{region 'Documentation'}
(*!
<summary>Capture once or compare against the retained snapshot after range validation.</summary>
*)
{endregion}
METHOD PROTECTED Assert
VAR
    ReferenceValue : REAL;
    ValuesEqual : BOOL;
    Value : REAL;
    InLowerIndex : DINT;
    InUpperIndex : DINT;
    MemoryLowerIndex : DINT;
    MemoryUpperIndex : DINT;
    MemoryEndIndex : LINT;
    EndIndex : LINT;
    Offset : LINT;
    InIndex : DINT;
    MemoryIndex : DINT;
    Message : STRING(GVL_Constants.MessageLength);
    ReferenceText : STRING(GVL_Constants.AssertionValueLength);
    ActualText : STRING(GVL_Constants.AssertionValueLength);
END_VAR
FEvaluationActive := ObservationActive AND FObservationPrevious AND FSnapshotValid;
FObservationPrevious := ObservationActive;

IF NOT ObservationActive THEN
    RETURN;
END_IF;

IF Result = E_Result.Error THEN
    RETURN;
END_IF;

// C0371: FB inputs are checked here before any reference access.
{warning disable C0371}
IF NOT __ISVALIDREF(IN) THEN
    Error(Message := 'Assertion error: IN reference is invalid.');
    RETURN;
END_IF;

IF NOT __ISVALIDREF(Memory) THEN
    Error(Message := 'Assertion error: Memory reference is invalid.');
    RETURN;
END_IF;

IF NOT Tc2_Utilities.RealIsFinite(x := Tolerance) THEN
    Error(Message := 'Assertion error: Tolerance must be finite.');
    RETURN;
END_IF;

IF Tolerance < 0.0 THEN
    Error(Message := 'Assertion error: Tolerance must not be negative.');
    RETURN;
END_IF;

InLowerIndex := LOWER_BOUND(IN, 1);
InUpperIndex := UPPER_BOUND(IN, 1);
MemoryLowerIndex := LOWER_BOUND(Memory, 1);
MemoryUpperIndex := UPPER_BOUND(Memory, 1);
EndIndex := DINT_TO_LINT(StartIndex) + USINT_TO_LINT(Length) - 1;
MemoryEndIndex := DINT_TO_LINT(MemoryLowerIndex) + USINT_TO_LINT(Length) - 1;

IF (Length = 0)
    OR (StartIndex < InLowerIndex) OR (StartIndex > InUpperIndex)
    OR (EndIndex > DINT_TO_LINT(InUpperIndex))
    OR (MemoryEndIndex > DINT_TO_LINT(MemoryUpperIndex)) THEN
    Message := CONCAT('Assertion error: array or memory range is invalid. StartIndex = ',
        DINT_TO_STRING(StartIndex));
    Message := CONCAT(Message, ', EndIndex = ');
    Message := CONCAT(Message, LINT_TO_STRING(EndIndex));
    Message := CONCAT(Message, ', Length = ');
    Message := CONCAT(Message, USINT_TO_STRING(Length));
    Message := CONCAT(Message, '.');
    Error(Message := Message);
    RETURN;
END_IF;

IF NOT FSnapshotValid THEN
    FOR Offset := 0 TO USINT_TO_LINT(Length) - 1 DO
        InIndex := LINT_TO_DINT(DINT_TO_LINT(StartIndex) + Offset);
        Value := IN[InIndex];
        IF Tc2_Utilities.RealIsNaN(x := Value) THEN
            Message := CONCAT('Assertion error: snapshot cannot contain NaN. IN index = ',
                DINT_TO_STRING(InIndex));
            Message := CONCAT(Message, '.');
            Error(Message := Message);
            RETURN;
        END_IF;
    END_FOR;
    FOR Offset := 0 TO USINT_TO_LINT(Length) - 1 DO
        InIndex := LINT_TO_DINT(DINT_TO_LINT(StartIndex) + Offset);
        MemoryIndex := LINT_TO_DINT(DINT_TO_LINT(MemoryLowerIndex) + Offset);
        Memory[MemoryIndex] := IN[InIndex];
    END_FOR;
    FSnapshotValid := TRUE;
    RETURN;
END_IF;

IF NOT EvaluationActive THEN
    RETURN;
END_IF;

IF Result = E_Result.Failed THEN
    RETURN;
END_IF;

FOR Offset := 0 TO USINT_TO_LINT(Length) - 1 DO
    InIndex := LINT_TO_DINT(DINT_TO_LINT(StartIndex) + Offset);
    MemoryIndex := LINT_TO_DINT(DINT_TO_LINT(MemoryLowerIndex) + Offset);
    Value := IN[InIndex];
    ReferenceValue := Memory[MemoryIndex];
    ValuesEqual := FALSE;
    IF NOT Tc2_Utilities.RealIsNaN(x := Value) THEN
        IF Value = ReferenceValue THEN
            ValuesEqual := TRUE;
        ELSIF Tc2_Utilities.RealIsFinite(x := Value)
            AND Tc2_Utilities.RealIsFinite(x := ReferenceValue) THEN
            ValuesEqual := IsWithinTolerance_Real(IN := Value,
                Expected := ReferenceValue,
                Tolerance := Tolerance);
        END_IF;
    END_IF;
    IF NOT ValuesEqual THEN
        Value := Memory[MemoryIndex];
        IF Tc2_Utilities.RealIsFinite(x := Value) THEN
            ReferenceText := CreateAssertionTextValue_Real(Value := Value);
        ELSE
            ReferenceText := '<non-finite>';
        END_IF;
        Value := IN[InIndex];
        IF Tc2_Utilities.RealIsFinite(x := Value) THEN
            ActualText := CreateAssertionTextValue_Real(Value := IN[InIndex]);
        ELSE
            ActualText := '<non-finite>';
        END_IF;
        Message := CONCAT('Assertion failed: array value changed. Reference[',
            DINT_TO_STRING(MemoryIndex));
        Message := CONCAT(Message, '] = ');
        Message := CONCAT(Message, ReferenceText);
        Message := CONCAT(Message, ', IN[');
        Message := CONCAT(Message, DINT_TO_STRING(InIndex));
        Message := CONCAT(Message, '] = ');
        Message := CONCAT(Message, ActualText);
        Message := CONCAT(Message, '.');
        Message := CONCAT(Message, ' Tolerance = ');
        Message := CONCAT(Message, CreateAssertionTextValue_Real(Value := Tolerance));
        Fail(Message := Message);
        RETURN;
    END_IF;
END_FOR;

Pass();
{warning restore C0371}
END_METHOD

{region 'Documentation'}
(*!
<summary>Current/last call has consecutive observation and an existing snapshot.</summary>
*)
{endregion}
{attribute 'monitoring' := 'call'}
PROPERTY PUBLIC EvaluationActive : BOOL //! Current/last call has consecutive observation and an existing snapshot.
GET // PUBLIC
EvaluationActive := FEvaluationActive;
END_GET
END_PROPERTY

{region 'Documentation'}
(*!
<summary>Invalidate the snapshot and observation history.</summary>
<description>

Does not clear external Memory. The next active observation captures a new snapshot
before comparison.

</description>
*)
{endregion}
METHOD PROTECTED ResetAssertion
FSnapshotValid := FALSE;
FObservationPrevious := FALSE;
FEvaluationActive := FALSE;
END_METHOD

END_FUNCTION_BLOCK

// ---- Framework/Assertions/POU/Utilities/IsWithinTolerance_Real.TcPOU
{region 'Documentation'}
(*!
<summary>Tests absolute tolerance without overflowing the typed difference. Requires finite inputs and a finite, non-negative tolerance; the caller validates them.</summary>
*)
{endregion}
FUNCTION INTERNAL IsWithinTolerance_Real : BOOL //! TRUE when the absolute difference is within Tolerance; caller must supply finite valid inputs.
VAR_INPUT
    IN : REAL; //! Actual value checked or observed by this Assertion.
    Expected : REAL; //! Reference value for comparison with IN.
    Tolerance : REAL; //! Maximum absolute difference accepted as equal; must be finite and non-negative.
END_VAR
VAR
    ActualMagnitude : REAL;
    ExpectedMagnitude : REAL;
    LargeMagnitude : REAL;
    SmallMagnitude : REAL;
    RemainingMagnitude : REAL;
    Difference : REAL;
END_VAR
VAR CONSTANT
    MaxFinite : REAL := REAL#3.40282346638528859811704183484516925440E38;
    HalfMaxFinite : REAL := MaxFinite / REAL#2.0;
END_VAR

IsWithinTolerance_Real := FALSE;

IF ((IN < 0.0) AND (Expected > 0.0)) OR ((IN > 0.0) AND (Expected < 0.0)) THEN
    ActualMagnitude := ABS(IN);
    ExpectedMagnitude := ABS(Expected);
    LargeMagnitude := MAX(ActualMagnitude, ExpectedMagnitude);
    SmallMagnitude := MIN(ActualMagnitude, ExpectedMagnitude);

    IF LargeMagnitude >= HalfMaxFinite THEN
        // Exact subtraction: MaxFinite and LargeMagnitude are within a factor of two.
        RemainingMagnitude := MaxFinite - LargeMagnitude;
        IF SmallMagnitude > RemainingMagnitude THEN
            RETURN;
        END_IF;
    END_IF;
END_IF;

Difference := ABS(IN - Expected);
IsWithinTolerance_Real := Difference <= Tolerance;

END_FUNCTION

// ---- Framework/Assertions/POU/Arrays/LReal/AssertArrayNoValueChange_LReal.TcPOU
{region 'Documentation'}
(*!
<summary>Captures one snapshot until Reset; Disable/Re-Enable never replaces it.</summary>
<description>

Disabling observation preserves the original snapshot. Re-enabling requires a fresh
preceding observation before comparisons resume; it does not replace that snapshot.

StartIndex is an absolute IN index and Length selects 1..255 elements within IN. Memory
must have at least Length elements from its own lower bound. Invalid references or ranges
report Error.

The caller provides dedicated writable Memory that must not overlap IN; overlap is not
checked. Keep bindings, selected range and snapshot contents stable until Reset. Reset
invalidates the snapshot without clearing Memory bytes.

Snapshot capture rejects NaN with Error but accepts either infinity. Later NaN is a
mismatch; equal signed infinities match.

Tolerance is absolute, in the same units as the values, finite and non-negative. Its
default zero requests exact comparison. The equality boundary is inclusive; larger differences
are unequal. Difference checking avoids overflow for large finite operands.

Numeric diagnostics use the formatter's default six significant digits; rounding affects
the message only, not the comparison.

</description>
*)
{endregion}
FUNCTION_BLOCK AssertArrayNoValueChange_LReal EXTENDS AssertionBase
VAR_INPUT
    Tolerance : LREAL := 0.0; //! Maximum absolute allowed difference; finite and non-negative.
    StartIndex : DINT; //! First selected index in IN; uses the array's declared index range, not a zero-based offset.
    Length : USINT; //! Number of monitored elements, from 1 through 255.
END_VAR
VAR_IN_OUT CONSTANT
    IN : ARRAY[*] OF LREAL; //! Read-only actual data; the selected range must remain stable during the call.
END_VAR
VAR_IN_OUT
    Memory : ARRAY[*] OF LREAL; //! Dedicated snapshot storage; only this assertion writes its selected elements.
END_VAR
VAR
    FSnapshotValid : BOOL;
    FObservationPrevious : BOOL;
    FEvaluationActive : BOOL;
END_VAR

SUPER^();

{region 'Documentation'}
(*!
<summary>Capture once or compare against the retained snapshot after range validation.</summary>
*)
{endregion}
METHOD PROTECTED Assert
VAR
    ReferenceValue : LREAL;
    ValuesEqual : BOOL;
    Value : LREAL;
    InLowerIndex : DINT;
    InUpperIndex : DINT;
    MemoryLowerIndex : DINT;
    MemoryUpperIndex : DINT;
    MemoryEndIndex : LINT;
    EndIndex : LINT;
    Offset : LINT;
    InIndex : DINT;
    MemoryIndex : DINT;
    Message : STRING(GVL_Constants.MessageLength);
    ReferenceText : STRING(GVL_Constants.AssertionValueLength);
    ActualText : STRING(GVL_Constants.AssertionValueLength);
END_VAR
FEvaluationActive := ObservationActive AND FObservationPrevious AND FSnapshotValid;
FObservationPrevious := ObservationActive;

IF NOT ObservationActive THEN
    RETURN;
END_IF;

IF Result = E_Result.Error THEN
    RETURN;
END_IF;

// C0371: FB inputs are checked here before any reference access.
{warning disable C0371}
IF NOT __ISVALIDREF(IN) THEN
    Error(Message := 'Assertion error: IN reference is invalid.');
    RETURN;
END_IF;

IF NOT __ISVALIDREF(Memory) THEN
    Error(Message := 'Assertion error: Memory reference is invalid.');
    RETURN;
END_IF;

IF NOT Tc2_Utilities.LrealIsFinite(x := Tolerance) THEN
    Error(Message := 'Assertion error: Tolerance must be finite.');
    RETURN;
END_IF;

IF Tolerance < 0.0 THEN
    Error(Message := 'Assertion error: Tolerance must not be negative.');
    RETURN;
END_IF;

InLowerIndex := LOWER_BOUND(IN, 1);
InUpperIndex := UPPER_BOUND(IN, 1);
MemoryLowerIndex := LOWER_BOUND(Memory, 1);
MemoryUpperIndex := UPPER_BOUND(Memory, 1);
EndIndex := DINT_TO_LINT(StartIndex) + USINT_TO_LINT(Length) - 1;
MemoryEndIndex := DINT_TO_LINT(MemoryLowerIndex) + USINT_TO_LINT(Length) - 1;

IF (Length = 0)
    OR (StartIndex < InLowerIndex) OR (StartIndex > InUpperIndex)
    OR (EndIndex > DINT_TO_LINT(InUpperIndex))
    OR (MemoryEndIndex > DINT_TO_LINT(MemoryUpperIndex)) THEN
    Message := CONCAT('Assertion error: array or memory range is invalid. StartIndex = ',
        DINT_TO_STRING(StartIndex));
    Message := CONCAT(Message, ', EndIndex = ');
    Message := CONCAT(Message, LINT_TO_STRING(EndIndex));
    Message := CONCAT(Message, ', Length = ');
    Message := CONCAT(Message, USINT_TO_STRING(Length));
    Message := CONCAT(Message, '.');
    Error(Message := Message);
    RETURN;
END_IF;

IF NOT FSnapshotValid THEN
    FOR Offset := 0 TO USINT_TO_LINT(Length) - 1 DO
        InIndex := LINT_TO_DINT(DINT_TO_LINT(StartIndex) + Offset);
        Value := IN[InIndex];
        IF Tc2_Utilities.LrealIsNaN(x := Value) THEN
            Message := CONCAT('Assertion error: snapshot cannot contain NaN. IN index = ',
                DINT_TO_STRING(InIndex));
            Message := CONCAT(Message, '.');
            Error(Message := Message);
            RETURN;
        END_IF;
    END_FOR;
    FOR Offset := 0 TO USINT_TO_LINT(Length) - 1 DO
        InIndex := LINT_TO_DINT(DINT_TO_LINT(StartIndex) + Offset);
        MemoryIndex := LINT_TO_DINT(DINT_TO_LINT(MemoryLowerIndex) + Offset);
        Memory[MemoryIndex] := IN[InIndex];
    END_FOR;
    FSnapshotValid := TRUE;
    RETURN;
END_IF;

IF NOT EvaluationActive THEN
    RETURN;
END_IF;

IF Result = E_Result.Failed THEN
    RETURN;
END_IF;

FOR Offset := 0 TO USINT_TO_LINT(Length) - 1 DO
    InIndex := LINT_TO_DINT(DINT_TO_LINT(StartIndex) + Offset);
    MemoryIndex := LINT_TO_DINT(DINT_TO_LINT(MemoryLowerIndex) + Offset);
    Value := IN[InIndex];
    ReferenceValue := Memory[MemoryIndex];
    ValuesEqual := FALSE;
    IF NOT Tc2_Utilities.LrealIsNaN(x := Value) THEN
        IF Value = ReferenceValue THEN
            ValuesEqual := TRUE;
        ELSIF Tc2_Utilities.LrealIsFinite(x := Value)
            AND Tc2_Utilities.LrealIsFinite(x := ReferenceValue) THEN
            ValuesEqual := IsWithinTolerance_LReal(IN := Value,
                Expected := ReferenceValue,
                Tolerance := Tolerance);
        END_IF;
    END_IF;
    IF NOT ValuesEqual THEN
        Value := Memory[MemoryIndex];
        IF Tc2_Utilities.LrealIsFinite(x := Value) THEN
            ReferenceText := CreateAssertionTextValue_LReal(Value := Value);
        ELSE
            ReferenceText := '<non-finite>';
        END_IF;
        Value := IN[InIndex];
        IF Tc2_Utilities.LrealIsFinite(x := Value) THEN
            ActualText := CreateAssertionTextValue_LReal(Value := IN[InIndex]);
        ELSE
            ActualText := '<non-finite>';
        END_IF;
        Message := CONCAT('Assertion failed: array value changed. Reference[',
            DINT_TO_STRING(MemoryIndex));
        Message := CONCAT(Message, '] = ');
        Message := CONCAT(Message, ReferenceText);
        Message := CONCAT(Message, ', IN[');
        Message := CONCAT(Message, DINT_TO_STRING(InIndex));
        Message := CONCAT(Message, '] = ');
        Message := CONCAT(Message, ActualText);
        Message := CONCAT(Message, '.');
        Message := CONCAT(Message, ' Tolerance = ');
        Message := CONCAT(Message, CreateAssertionTextValue_LReal(Value := Tolerance));
        Fail(Message := Message);
        RETURN;
    END_IF;
END_FOR;

Pass();
{warning restore C0371}
END_METHOD

{region 'Documentation'}
(*!
<summary>Current/last call has consecutive observation and an existing snapshot.</summary>
*)
{endregion}
{attribute 'monitoring' := 'call'}
PROPERTY PUBLIC EvaluationActive : BOOL //! Current/last call has consecutive observation and an existing snapshot.
GET // PUBLIC
EvaluationActive := FEvaluationActive;
END_GET
END_PROPERTY

{region 'Documentation'}
(*!
<summary>Invalidate the snapshot and observation history.</summary>
<description>

Does not clear external Memory. The next active observation captures a new snapshot
before comparison.

</description>
*)
{endregion}
METHOD PROTECTED ResetAssertion
FSnapshotValid := FALSE;
FObservationPrevious := FALSE;
FEvaluationActive := FALSE;
END_METHOD

END_FUNCTION_BLOCK

// ---- SelfTests/TestSuites/TestSuite_AssertionText.TcPOU
{region 'Documentation'}
(*!
<summary>Checks text, token and diagnostic boundaries with isolated Assertion subjects.</summary>
*)
{endregion}
FUNCTION_BLOCK TestSuite_AssertionText EXTENDS TestSuiteBase
VAR
    FTextComparison : Test_AssertionTextComparison;
    FTextSearch : Test_AssertionTextSearch;
    FTextDiagnostics : Test_AssertionTextDiagnostics;
    FValueTokenCount : Test_AssertionValueTokenCount;
    FArrayTokenCount : Test_AssertionArrayTokenCount;
    FLengthUntil : Test_AssertionLengthUntil;
    FTestCases : ARRAY[1..TestCaseCapacity] OF I_TestCase;
END_VAR
VAR CONSTANT
    TestCaseCapacity : UINT := 6;
END_VAR

SUPER^();

{region 'Documentation'}
(*!
<summary>Initializes six isolated text and token Test Cases and registers them serially.</summary>
*)
{endregion}
METHOD PROTECTED Configure
VAR_IN_OUT
    // SA0167: Borrowed owner builder; no temporary instance is created.
    {attribute 'analysis' := '-167'}
    Builder : TestSuiteConfigurationBuilder; //! Borrowed owner configuration builder used only during this Configure call; register this owner's concrete children.
END_VAR
VAR
    TestConfig : ST_TestCaseConfig;
END_VAR
Builder.Initialize(Mode := E_OrchestrationMode.Serial,
    TestCases := FTestCases);
FTextComparison.Initialize(Parent := THIS^,
    TestName := 'TextComparison',
    Config := TestConfig);
Builder.Register(TestCase := FTextComparison);
FTextSearch.Initialize(Parent := THIS^,
    TestName := 'TextSearch',
    Config := TestConfig);
Builder.Register(TestCase := FTextSearch);
FTextDiagnostics.Initialize(Parent := THIS^,
    TestName := 'TextDiagnostics',
    Config := TestConfig);
Builder.Register(TestCase := FTextDiagnostics);
FValueTokenCount.Initialize(Parent := THIS^,
    TestName := 'ValueTokenCount',
    Config := TestConfig);
Builder.Register(TestCase := FValueTokenCount);
FArrayTokenCount.Initialize(Parent := THIS^,
    TestName := 'ArrayTokenCount',
    Config := TestConfig);
Builder.Register(TestCase := FArrayTokenCount);
FLengthUntil.Initialize(Parent := THIS^,
    TestName := 'LengthUntil',
    Config := TestConfig);
Builder.Register(TestCase := FLengthUntil);
END_METHOD

{region 'Documentation'}
(*!
<summary>Returns a registered scenario using its original array index.</summary>
*)
{endregion}
METHOD PUBLIC GetTestCase : I_TestCase //! Typed child interface at the original array index; zero when no entry is available.
VAR_INPUT
    Index : DINT; //! Original occupied child-array index, rather than an ordinal position.
END_VAR
GetTestCase := 0;
IF (ChildCount = 0) OR (Index < ChildArrayLowerBound)
    OR (DINT_TO_LINT(Index) >= DINT_TO_LINT(ChildArrayLowerBound) + UINT_TO_LINT(ChildCount)) THEN
    RETURN;
END_IF;
GetTestCase := FTestCases[Index];
END_METHOD

{region 'Documentation'}
(*!
<summary>Calls every owned scenario once per initialized Suite cycle.</summary>
*)
{endregion}
METHOD PROTECTED ProcessTestCases
FTextComparison();
FTextSearch();
FTextDiagnostics();
FValueTokenCount();
FArrayTokenCount();
FLengthUntil();
END_METHOD

END_FUNCTION_BLOCK

// ---- SelfTests/TestCases/TestSuite_AssertionText/Test_AssertionTextComparison.TcPOU
{region 'Documentation'}
(*!
<summary>Checks exact STRING/WSTRING comparisons and configured length boundaries.</summary>
<description>
Equality and inequality share explicit operands, but each result is asserted.
Wide-code-unit cases distinguish a zero low byte from the WSTRING terminator
and equal low bytes from equal code units. Capacity tests use the configured
content limits, including the last character and one excessive character.
Each scenario occupies two calls: Reset with valid bindings, then evaluation.
ProcessAssertions checks each call before ProcessTests advances. Literal expected
results belong to SelectScenario, not to a copy of the production comparison.
The local capture is cleared before each call and checked in subject-call order.
FirstFailedScenario and FailedDuringEvaluation retain the first mismatch.
Caller text buffers provide at least one extra character of capacity so overlength tests
reach the real read-only reference API without an intermediate truncating copy.
</description>
*)
{endregion}
FUNCTION_BLOCK Test_AssertionTextComparison EXTENDS TestCaseBase
VAR
    FEqual : AssertEqual_String;
    FEqualExpectedResult : E_Result;
    FNotEqual : AssertNotEqual_String;
    FNotEqualExpectedResult : E_Result;
    FWideEqual : AssertEqual_WString;
    FWideEqualExpectedResult : E_Result;
    FWideNotEqual : AssertNotEqual_WString;
    FWideNotEqualExpectedResult : E_Result;
    FInput : STRING(InputCapacity);
    FInputBefore : STRING(InputCapacity);
    FWideInput : WSTRING(WideInputCapacity);
    FWideInputBefore : WSTRING(WideInputCapacity);
    FExpected : STRING(InputCapacity);
    FExpectedBefore : STRING(InputCapacity);
    FWideExpected : WSTRING(WideInputCapacity);
    FWideExpectedBefore : WSTRING(WideInputCapacity);
    FCapture : EventBuffer;
    FEvents : ARRAY[1..CaptureLength] OF ST_Event;
    FCaptureFifo : ST_FifoStatus;
    FCaptureStatus : ST_EventBufferStatus;
    FSetupValid : BOOL;
    FScenario : UINT;
    FChecked : BOOL;
    FEvaluateSubjects : BOOL;
    FObservationReady : BOOL;
    FFirstFailedScenario : UINT;
    FFailedDuringEvaluation : BOOL;
    FResultsMatch : BOOL;
    FResults : AssertTrue;
    FActivityMatch : BOOL;
    FActivity : AssertTrue;
    FInputsMatch : BOOL;
    FInputs : AssertTrue;
    FFindingsMatch : BOOL;
    FFindings : AssertTrue;
END_VAR
VAR CONSTANT
    InputCapacity : UINT := Param_Assertions.AssertionStringLength + 1;
    // XAE rejects a computed WSTRING capacity here. Covers the default limit plus one.
    // CheckInitialization rejects a configuration exceeding this test storage.
    WideInputCapacity : UINT := 81;
    CaptureLength : UINT := 8;
    ScenarioExact : UINT := 1;
    ScenarioEmpty : UINT := 2;
    ScenarioCaseSensitive : UINT := 3;
    ScenarioFirstCharacter : UINT := 4;
    ScenarioLastCharacter : UINT := 5;
    ScenarioDifferentLength : UINT := 6;
    ScenarioWideHighByte : UINT := 7;
    ScenarioWideZeroLowByte : UINT := 8;
    ScenarioBelowCapacity : UINT := 9;
    ScenarioAtCapacity : UINT := 10;
    ScenarioLastAtCapacity : UINT := 11;
    ScenarioInputOverCapacity : UINT := 12;
    ScenarioExpectedOverCapacity : UINT := 13;
    LastScenario : UINT := ScenarioExpectedOverCapacity;
END_VAR

SUPER^();

{region 'Documentation'}
(*!
<summary>Aggregates only outer checks, not intentionally failing subjects.</summary>
*)
{endregion}
METHOD PROTECTED AggregateResults
VAR_INPUT
    Aggregator : I_ResultAggregator; //! Borrowed result sink owned by the outer Test Case; add this test's checking Assertions without resetting or retaining the sink.
END_VAR
Aggregator.AddProvider(Provider := FResults);
Aggregator.AddProvider(Provider := FActivity);
Aggregator.AddProvider(Provider := FInputs);
Aggregator.AddProvider(Provider := FFindings);
END_METHOD

{region 'Documentation'}
(*!
<summary>Calls each inherited production subject once with caller-owned text storage.</summary>
*)
{endregion}
METHOD PRIVATE CallSubjects
FEqual(Enable := TRUE,
    State := E_State.Running,
    IN := FInput,
    Expected := FExpected);
FNotEqual(Enable := TRUE,
    State := E_State.Running,
    IN := FInput,
    Expected := FExpected);
FWideEqual(Enable := TRUE,
    State := E_State.Running,
    IN := FWideInput,
    Expected := FWideExpected);
FWideNotEqual(Enable := TRUE,
    State := E_State.Running,
    IN := FWideInput,
    Expected := FWideExpected);
END_METHOD

{region 'Documentation'}
(*!
<summary>Checks one subject finding in call order; expected outcomes come from the scenario.</summary>
*)
{endregion}
METHOD PRIVATE CheckFinding : BOOL //! TRUE when the required finding checks pass; calls requiring no finding also succeed.
VAR_INPUT
    Subject : I_Assertion; //! Assertion interface supplying the expected finding identity.
    ExpectedResult : E_Result; //! Independently authored result expected in the captured finding.
END_VAR
VAR_IN_OUT
    Index : UINT; //! One-based next finding index; advanced when this call checks a required finding.
END_VAR
CheckFinding := TRUE;
IF FEvaluateSubjects AND ((ExpectedResult = E_Result.Failed)
    OR (ExpectedResult = E_Result.Error)) THEN
    CheckFinding := (FEvents[Index].SequenceId = UINT_TO_UDINT(Index))
        AND (FEvents[Index].Name = Subject.Name)
        AND (FEvents[Index].OwnerScope = E_OwnerScope.Assertion)
        AND (FEvents[Index].EventType = E_EventType.Result)
        AND (FEvents[Index].State = E_State.Running)
        AND (FEvents[Index].Result = ExpectedResult)
        AND (FEvents[Index].Message <> '');
    Index := Index + 1;
END_IF;
END_METHOD

{region 'Documentation'}
(*!
<summary>Checks exact finding count and identities; at most one finding per subject.</summary>
*)
{endregion}
METHOD PRIVATE CheckFindings
VAR
    Index : UINT;
    Matches : BOOL;
END_VAR
Index := 1;
FFindingsMatch := TRUE;
Matches := CheckFinding(Subject := FEqual,
    ExpectedResult := FEqualExpectedResult,
    Index := Index);
FFindingsMatch := FFindingsMatch AND Matches;
Matches := CheckFinding(Subject := FNotEqual,
    ExpectedResult := FNotEqualExpectedResult,
    Index := Index);
FFindingsMatch := FFindingsMatch AND Matches;
Matches := CheckFinding(Subject := FWideEqual,
    ExpectedResult := FWideEqualExpectedResult,
    Index := Index);
FFindingsMatch := FFindingsMatch AND Matches;
Matches := CheckFinding(Subject := FWideNotEqual,
    ExpectedResult := FWideNotEqualExpectedResult,
    Index := Index);
FFindingsMatch := FFindingsMatch AND Matches;
FFindingsMatch := FFindingsMatch
    AND (FCaptureStatus.SequenceId = UINT_TO_UDINT(Index - 1))
    AND (FCaptureStatus.LostEventCount = 0);
END_METHOD

{region 'Documentation'}
(*!
<summary>Rejects incomplete subject, capture or outer Assertion setup.</summary>
*)
{endregion}
METHOD PROTECTED CheckInitialization : BOOL //! TRUE when the inherited initialization check and this concrete fixture check both accept the setup.
CheckInitialization := SUPER^.CheckInitialization();
IF NOT CheckInitialization THEN
    RETURN;
END_IF;

CheckInitialization := FSetupValid
    AND (Param_Assertions.AssertionStringLength >= 5)
    AND (Param_Assertions.AssertionWStringLength >= 5)
    AND (Param_Assertions.AssertionWStringLength < WideInputCapacity)
    AND FResults.IsInitialized
    AND FActivity.IsInitialized
    AND FInputs.IsInitialized
    AND FFindings.IsInitialized;
IF NOT CheckInitialization THEN
    EventPublisher.PublishEvent(Event := CreateFrameworkEvent(Name := Name,
        ResourceName := '',
        State := State,
        Severity := E_EventSeverity.Error,
        Message := 'Text selftest setup failed.'));
END_IF;
END_METHOD

{region 'Documentation'}
(*!
<summary>Checks literal evaluation results, or NotEvaluated on the reset call.</summary>
*)
{endregion}
METHOD PRIVATE CheckResults
IF FEvaluateSubjects THEN
    FResultsMatch := (FEqual.Result = FEqualExpectedResult)
        AND (FNotEqual.Result = FNotEqualExpectedResult)
        AND (FWideEqual.Result = FWideEqualExpectedResult)
        AND (FWideNotEqual.Result = FWideNotEqualExpectedResult);
ELSE
    FResultsMatch := (FEqual.Result = E_Result.NotEvaluated)
        AND (FNotEqual.Result = E_Result.NotEvaluated)
        AND (FWideEqual.Result = E_Result.NotEvaluated)
        AND (FWideNotEqual.Result = E_Result.NotEvaluated);
END_IF;
FActivityMatch := FEqual.Enabled
    AND (FEqual.ObservationActive = FEvaluateSubjects)
    AND (FEqual.EvaluationActive = FEvaluateSubjects)
    AND FNotEqual.Enabled
    AND (FNotEqual.ObservationActive = FEvaluateSubjects)
    AND (FNotEqual.EvaluationActive = FEvaluateSubjects)
    AND FWideEqual.Enabled
    AND (FWideEqual.ObservationActive = FEvaluateSubjects)
    AND (FWideEqual.EvaluationActive = FEvaluateSubjects)
    AND FWideNotEqual.Enabled
    AND (FWideNotEqual.ObservationActive = FEvaluateSubjects)
    AND (FWideNotEqual.EvaluationActive = FEvaluateSubjects);
END_METHOD

{region 'Documentation'}
(*!
<summary>Initializes outer checks and isolates intentional subject findings.</summary>
*)
{endregion}
METHOD PROTECTED Configure
VAR
    Initialized : BOOL;
END_VAR
FPreparationStateCount := 0;
FTestStateCount := 1;
FResults.Initialize(Parent := THIS^,
    AssertionName := 'Results');
FActivity.Initialize(Parent := THIS^,
    AssertionName := 'Activity');
FInputs.Initialize(Parent := THIS^,
    AssertionName := 'Inputs');
FFindings.Initialize(Parent := THIS^,
    AssertionName := 'Findings');
FSetupValid := FCapture.Initialize(Buffer := FEvents,
    FifoControl := FCaptureFifo,
    Status := FCaptureStatus);
FEqual.BindPublisher(Publisher := FCapture);
Initialized := FEqual.Initialize(Parent := THIS^,
    AssertionName := 'Equal');
FSetupValid := FSetupValid AND Initialized;
FNotEqual.BindPublisher(Publisher := FCapture);
Initialized := FNotEqual.Initialize(Parent := THIS^,
    AssertionName := 'NotEqual');
FSetupValid := FSetupValid AND Initialized;
FWideEqual.BindPublisher(Publisher := FCapture);
Initialized := FWideEqual.Initialize(Parent := THIS^,
    AssertionName := 'WideEqual');
FSetupValid := FSetupValid AND Initialized;
FWideNotEqual.BindPublisher(Publisher := FCapture);
Initialized := FWideNotEqual.Initialize(Parent := THIS^,
    AssertionName := 'WideNotEqual');
FSetupValid := FSetupValid AND Initialized;
END_METHOD

{region 'Documentation'}
(*!
<summary>Completes abort; no asynchronous resource is owned.</summary>
*)
{endregion}
METHOD PROTECTED ProcessAbort
VAR_INPUT
    Enable : BOOL; //! Phase permission supplied by the owning Test Case; FALSE does not authorize progression, while observation may continue.
END_VAR
IF Enable THEN
    CompleteAbort();
END_IF;
END_METHOD

{region 'Documentation'}
(*!
<summary>Latches this call's checks before progression is permitted.</summary>
*)
{endregion}
METHOD PROTECTED ProcessAssertions
VAR_INPUT
    Enable : BOOL; //! Phase permission supplied by the owning Test Case; FALSE does not authorize progression, while observation may continue.
END_VAR
VAR
    Check : BOOL;
END_VAR
Check := Enable AND FObservationReady;
FResults(Enable := Check,
    State := State,
    IN := FResultsMatch);
FActivity(Enable := Check,
    State := State,
    IN := FActivityMatch);
FInputs(Enable := Check,
    State := State,
    IN := FInputsMatch);
FFindings(Enable := Check,
    State := State,
    IN := FFindingsMatch);
IF Check THEN
    FChecked := TRUE;
END_IF;
END_METHOD

{region 'Documentation'}
(*!
<summary>No Preparation phase is needed.</summary>
*)
{endregion}
METHOD PROTECTED ProcessPreparations
VAR_INPUT
    // SA0033: Required hook; this test has no Preparation phase.
    {attribute 'analysis' := '-33'}
    Enable : BOOL; //! Phase permission supplied by the owning Test Case; FALSE does not authorize progression, while observation may continue.
END_VAR
END_METHOD

{region 'Documentation'}
(*!
<summary>Restarts the scenario sequence and outer checks.</summary>
*)
{endregion}
METHOD PROTECTED ProcessReset
FScenario := ScenarioExact;
FChecked := FALSE;
FEvaluateSubjects := FALSE;
FObservationReady := FALSE;
FFirstFailedScenario := 0;
FFailedDuringEvaluation := FALSE;
FCapture.Reset();
ResetSubjects();
FResults.Reset();
FActivity.Reset();
FInputs.Reset();
FFindings.Reset();
CompleteReset();
END_METHOD

{region 'Documentation'}
(*!
<summary>Resets then evaluates each scenario on separate cycles before advancing.</summary>
*)
{endregion}
METHOD PROTECTED ProcessTests
VAR_INPUT
    Enable : BOOL; //! Phase permission supplied by the owning Test Case; FALSE does not authorize progression, while observation may continue.
END_VAR
IF NOT Enable THEN
    RETURN;
END_IF;

IF FChecked THEN
    FChecked := FALSE;
    FObservationReady := FALSE;
    IF FEvaluateSubjects THEN
        IF FScenario = LastScenario THEN
            CompleteTests();
            RETURN;
        END_IF;
        FScenario := FScenario + 1;
    END_IF;
    FEvaluateSubjects := NOT FEvaluateSubjects;
END_IF;

IF NOT SelectScenario() THEN
    RETURN;
END_IF;
FCapture.Reset();
IF NOT FEvaluateSubjects THEN
    ResetSubjects();
END_IF;
FInputBefore := FInput;
FWideInputBefore := FWideInput;
FExpectedBefore := FExpected;
FWideExpectedBefore := FWideExpected;
CallSubjects();
CheckResults();
FInputsMatch := (FInput = FInputBefore)
    AND (FWideInput = FWideInputBefore)
    AND (FExpected = FExpectedBefore)
    AND (FWideExpected = FWideExpectedBefore);
CheckFindings();
IF (FFirstFailedScenario = 0)
    AND NOT (FResultsMatch AND FActivityMatch AND FInputsMatch AND FFindingsMatch) THEN
    FFirstFailedScenario := FScenario;
    FFailedDuringEvaluation := FEvaluateSubjects;
END_IF;
FObservationReady := TRUE;
END_METHOD

{region 'Documentation'}
(*!
<summary>Queues reset; the next bound FB call consumes it without evaluating.</summary>
*)
{endregion}
METHOD PRIVATE ResetSubjects
FEqual.Reset();
FNotEqual.Reset();
FWideEqual.Reset();
FWideNotEqual.Reset();
END_METHOD

{region 'Documentation'}
(*!
<summary>Selects explicit text stimuli and expected results for one scenario.</summary>
*)
{endregion}
METHOD PRIVATE SelectScenario : BOOL //! TRUE after selecting a supported scenario and its literal expectations; FALSE reports an unknown scenario.
VAR
    Index : UINT;
END_VAR
SelectScenario := FALSE;
FInput := 'ABC';
FExpected := 'ABC';
FWideInput := "ABC";
FWideExpected := "ABC";
CASE FScenario OF
    ScenarioExact:

        FEqualExpectedResult := E_Result.Passed;
        FNotEqualExpectedResult := E_Result.Failed;
        FWideEqualExpectedResult := E_Result.Passed;
        FWideNotEqualExpectedResult := E_Result.Failed;
    ScenarioEmpty:
        FInput := '';
        FExpected := '';
        FWideInput := "";
        FWideExpected := "";
        FEqualExpectedResult := E_Result.Passed;
        FNotEqualExpectedResult := E_Result.Failed;
        FWideEqualExpectedResult := E_Result.Passed;
        FWideNotEqualExpectedResult := E_Result.Failed;
    ScenarioCaseSensitive:
        FExpected := 'AbC';
        FWideExpected := "AbC";
        FEqualExpectedResult := E_Result.Failed;
        FNotEqualExpectedResult := E_Result.Passed;
        FWideEqualExpectedResult := E_Result.Failed;
        FWideNotEqualExpectedResult := E_Result.Passed;
    ScenarioFirstCharacter:
        FExpected := 'ZBC';
        FWideExpected := "ZBC";
        FEqualExpectedResult := E_Result.Failed;
        FNotEqualExpectedResult := E_Result.Passed;
        FWideEqualExpectedResult := E_Result.Failed;
        FWideNotEqualExpectedResult := E_Result.Passed;
    ScenarioLastCharacter:
        FExpected := 'ABZ';
        FWideExpected := "ABZ";
        FEqualExpectedResult := E_Result.Failed;
        FNotEqualExpectedResult := E_Result.Passed;
        FWideEqualExpectedResult := E_Result.Failed;
        FWideNotEqualExpectedResult := E_Result.Passed;
    ScenarioDifferentLength:
        FExpected := 'AB';
        FWideExpected := "AB";
        FEqualExpectedResult := E_Result.Failed;
        FNotEqualExpectedResult := E_Result.Passed;
        FWideEqualExpectedResult := E_Result.Failed;
        FWideNotEqualExpectedResult := E_Result.Passed;
    ScenarioWideHighByte:
        FWideInput[0] := WORD#16#0141;
        FWideExpected[0] := WORD#16#0241;
        FEqualExpectedResult := E_Result.Passed;
        FNotEqualExpectedResult := E_Result.Failed;
        FWideEqualExpectedResult := E_Result.Failed;
        FWideNotEqualExpectedResult := E_Result.Passed;
    ScenarioWideZeroLowByte:
        FWideInput[0] := WORD#16#0100;
        FWideExpected[0] := WORD#16#0100;
        FWideExpected[2] := WORD#16#005A;
        FEqualExpectedResult := E_Result.Passed;
        FNotEqualExpectedResult := E_Result.Failed;
        FWideEqualExpectedResult := E_Result.Failed;
        FWideNotEqualExpectedResult := E_Result.Passed;
    ScenarioBelowCapacity:
        FOR Index := 0 TO Param_Assertions.AssertionStringLength DO
            // SA0175: Bounded byte writes construct exact input/terminator boundaries; no UTF-8 decoding.
            {analysis -175}
            FInput[Index] := BYTE#16#41;
            FExpected[Index] := BYTE#16#41;
            {analysis +175}
        END_FOR;
        // SA0175: Bounded byte writes construct exact input/terminator boundaries; no UTF-8 decoding.
        {analysis -175}
        FInput[Param_Assertions.AssertionStringLength - 1] := 0;
        FExpected[Param_Assertions.AssertionStringLength - 1] := 0;
        {analysis +175}
        FOR Index := 0 TO Param_Assertions.AssertionWStringLength DO
            FWideInput[Index] := WORD#16#0141;
            FWideExpected[Index] := WORD#16#0141;
        END_FOR;
        FWideInput[Param_Assertions.AssertionWStringLength - 1] := 0;
        FWideExpected[Param_Assertions.AssertionWStringLength - 1] := 0;
        FEqualExpectedResult := E_Result.Passed;
        FNotEqualExpectedResult := E_Result.Failed;
        FWideEqualExpectedResult := E_Result.Passed;
        FWideNotEqualExpectedResult := E_Result.Failed;
    ScenarioAtCapacity:
        FOR Index := 0 TO Param_Assertions.AssertionStringLength DO
            // SA0175: Bounded byte writes construct exact input/terminator boundaries; no UTF-8 decoding.
            {analysis -175}
            FInput[Index] := BYTE#16#41;
            FExpected[Index] := BYTE#16#41;
            {analysis +175}
        END_FOR;
        // SA0175: Bounded byte writes construct exact input/terminator boundaries; no UTF-8 decoding.
        {analysis -175}
        FInput[Param_Assertions.AssertionStringLength] := 0;
        FExpected[Param_Assertions.AssertionStringLength] := 0;
        {analysis +175}
        FOR Index := 0 TO Param_Assertions.AssertionWStringLength DO
            FWideInput[Index] := WORD#16#0141;
            FWideExpected[Index] := WORD#16#0141;
        END_FOR;
        FWideInput[Param_Assertions.AssertionWStringLength] := 0;
        FWideExpected[Param_Assertions.AssertionWStringLength] := 0;
        FEqualExpectedResult := E_Result.Passed;
        FNotEqualExpectedResult := E_Result.Failed;
        FWideEqualExpectedResult := E_Result.Passed;
        FWideNotEqualExpectedResult := E_Result.Failed;
    ScenarioLastAtCapacity:
        FOR Index := 0 TO Param_Assertions.AssertionStringLength DO
            // SA0175: Bounded byte writes construct exact input/terminator boundaries; no UTF-8 decoding.
            {analysis -175}
            FInput[Index] := BYTE#16#41;
            FExpected[Index] := BYTE#16#41;
            {analysis +175}
        END_FOR;
        // SA0175: Bounded byte writes construct exact input/terminator boundaries; no UTF-8 decoding.
        {analysis -175}
        FInput[Param_Assertions.AssertionStringLength] := 0;
        FExpected[Param_Assertions.AssertionStringLength] := 0;
        {analysis +175}
        FOR Index := 0 TO Param_Assertions.AssertionWStringLength DO
            FWideInput[Index] := WORD#16#0141;
            FWideExpected[Index] := WORD#16#0141;
        END_FOR;
        FWideInput[Param_Assertions.AssertionWStringLength] := 0;
        FWideExpected[Param_Assertions.AssertionWStringLength] := 0;
        // SA0175: Bounded byte writes construct exact input/terminator boundaries; no UTF-8 decoding.
        {analysis -175}
        FExpected[Param_Assertions.AssertionStringLength - 1] := BYTE#16#42;
        {analysis +175}
        FWideExpected[Param_Assertions.AssertionWStringLength - 1] := WORD#16#0241;
        FEqualExpectedResult := E_Result.Failed;
        FNotEqualExpectedResult := E_Result.Passed;
        FWideEqualExpectedResult := E_Result.Failed;
        FWideNotEqualExpectedResult := E_Result.Passed;
    ScenarioInputOverCapacity:
        FOR Index := 0 TO Param_Assertions.AssertionStringLength DO
            // SA0175: Bounded byte writes construct exact input/terminator boundaries; no UTF-8 decoding.
            {analysis -175}
            FInput[Index] := BYTE#16#41;
            FExpected[Index] := BYTE#16#41;
            {analysis +175}
        END_FOR;
        // SA0175: Bounded byte writes construct exact input/terminator boundaries; no UTF-8 decoding.
        {analysis -175}
        FInput[Param_Assertions.AssertionStringLength] := 0;
        FExpected[Param_Assertions.AssertionStringLength] := 0;
        {analysis +175}
        FOR Index := 0 TO Param_Assertions.AssertionWStringLength DO
            FWideInput[Index] := WORD#16#0141;
            FWideExpected[Index] := WORD#16#0141;
        END_FOR;
        FWideInput[Param_Assertions.AssertionWStringLength] := 0;
        FWideExpected[Param_Assertions.AssertionWStringLength] := 0;
        // SA0175: Bounded byte writes construct exact input/terminator boundaries; no UTF-8 decoding.
        {analysis -175}
        FInput[Param_Assertions.AssertionStringLength] := BYTE#16#41;
        FInput[Param_Assertions.AssertionStringLength + 1] := 0;
        {analysis +175}
        FWideInput[Param_Assertions.AssertionWStringLength] := WORD#16#0141;
        FWideInput[Param_Assertions.AssertionWStringLength + 1] := 0;
        FEqualExpectedResult := E_Result.Error;
        FNotEqualExpectedResult := E_Result.Error;
        FWideEqualExpectedResult := E_Result.Error;
        FWideNotEqualExpectedResult := E_Result.Error;
    ScenarioExpectedOverCapacity:
        FOR Index := 0 TO Param_Assertions.AssertionStringLength DO
            // SA0175: Bounded byte writes construct exact input/terminator boundaries; no UTF-8 decoding.
            {analysis -175}
            FInput[Index] := BYTE#16#41;
            FExpected[Index] := BYTE#16#41;
            {analysis +175}
        END_FOR;
        // SA0175: Bounded byte writes construct exact input/terminator boundaries; no UTF-8 decoding.
        {analysis -175}
        FInput[Param_Assertions.AssertionStringLength] := 0;
        FExpected[Param_Assertions.AssertionStringLength] := 0;
        {analysis +175}
        FOR Index := 0 TO Param_Assertions.AssertionWStringLength DO
            FWideInput[Index] := WORD#16#0141;
            FWideExpected[Index] := WORD#16#0141;
        END_FOR;
        FWideInput[Param_Assertions.AssertionWStringLength] := 0;
        FWideExpected[Param_Assertions.AssertionWStringLength] := 0;
        // SA0175: Bounded byte writes construct exact input/terminator boundaries; no UTF-8 decoding.
        {analysis -175}
        FExpected[Param_Assertions.AssertionStringLength] := BYTE#16#41;
        FExpected[Param_Assertions.AssertionStringLength + 1] := 0;
        {analysis +175}
        FWideExpected[Param_Assertions.AssertionWStringLength] := WORD#16#0141;
        FWideExpected[Param_Assertions.AssertionWStringLength + 1] := 0;
        FEqualExpectedResult := E_Result.Error;
        FNotEqualExpectedResult := E_Result.Error;
        FWideEqualExpectedResult := E_Result.Error;
        FWideNotEqualExpectedResult := E_Result.Error;
ELSE
    Error(Message := 'Unknown text scenario.');
    RETURN;
END_CASE;
SelectScenario := TRUE;
END_METHOD

END_FUNCTION_BLOCK

// ---- SelfTests/TestCases/TestSuite_AssertionText/Test_AssertionTextSearch.TcPOU
{region 'Documentation'}
(*!
<summary>Checks prefix, suffix and containment with bounded STRING/WSTRING inputs.</summary>
<description>
Explicit vectors cover first/last candidates, whole input, absent and longer
fragments, empty-input Failed versus empty-fragment Error, and maximum content.
Wide text includes nonzero code units with a zero low byte and high-byte-only
differences. Matching is exact and case-sensitive; no text normalization is used.
Each scenario occupies two calls: Reset with valid bindings, then evaluation.
ProcessAssertions checks each call before ProcessTests advances. Literal expected
results belong to SelectScenario, not to a copy of the production comparison.
The local capture is cleared before each call and checked in subject-call order.
FirstFailedScenario and FailedDuringEvaluation retain the first mismatch.
Caller text buffers provide at least one extra character of capacity so overlength tests
reach the real read-only reference API without an intermediate truncating copy.
</description>
*)
{endregion}
FUNCTION_BLOCK Test_AssertionTextSearch EXTENDS TestCaseBase
VAR
    FStartsWith : AssertStartsWith_String;
    FStartsWithExpectedResult : E_Result;
    FEndsWith : AssertEndsWith_String;
    FEndsWithExpectedResult : E_Result;
    FContains : AssertContains_String;
    FContainsExpectedResult : E_Result;
    FWideStartsWith : AssertStartsWith_WString;
    FWideStartsWithExpectedResult : E_Result;
    FWideEndsWith : AssertEndsWith_WString;
    FWideEndsWithExpectedResult : E_Result;
    FWideContains : AssertContains_WString;
    FWideContainsExpectedResult : E_Result;
    FInput : STRING(InputCapacity);
    FInputBefore : STRING(InputCapacity);
    FWideInput : WSTRING(WideInputCapacity);
    FWideInputBefore : WSTRING(WideInputCapacity);
    FPrefix : STRING(InputCapacity);
    FPrefixBefore : STRING(InputCapacity);
    FWidePrefix : WSTRING(WideInputCapacity);
    FWidePrefixBefore : WSTRING(WideInputCapacity);
    FSuffix : STRING(InputCapacity);
    FSuffixBefore : STRING(InputCapacity);
    FWideSuffix : WSTRING(WideInputCapacity);
    FWideSuffixBefore : WSTRING(WideInputCapacity);
    FFragment : STRING(InputCapacity);
    FFragmentBefore : STRING(InputCapacity);
    FWideFragment : WSTRING(WideInputCapacity);
    FWideFragmentBefore : WSTRING(WideInputCapacity);
    FCapture : EventBuffer;
    FEvents : ARRAY[1..CaptureLength] OF ST_Event;
    FCaptureFifo : ST_FifoStatus;
    FCaptureStatus : ST_EventBufferStatus;
    FSetupValid : BOOL;
    FScenario : UINT;
    FChecked : BOOL;
    FEvaluateSubjects : BOOL;
    FObservationReady : BOOL;
    FFirstFailedScenario : UINT;
    FFailedDuringEvaluation : BOOL;
    FResultsMatch : BOOL;
    FResults : AssertTrue;
    FActivityMatch : BOOL;
    FActivity : AssertTrue;
    FInputsMatch : BOOL;
    FInputs : AssertTrue;
    FFindingsMatch : BOOL;
    FFindings : AssertTrue;
END_VAR
VAR CONSTANT
    InputCapacity : UINT := Param_Assertions.AssertionStringLength + 1;
    // XAE rejects a computed WSTRING capacity here. Covers the default limit plus one.
    // CheckInitialization rejects a configuration exceeding this test storage.
    WideInputCapacity : UINT := 81;
    // Six findings must remain below the buffer's Length - 2 diagnostic threshold.
    CaptureLength : UINT := 10;
    ScenarioMatching : UINT := 1;
    ScenarioWholeInput : UINT := 2;
    ScenarioFirstPosition : UINT := 3;
    ScenarioLastPosition : UINT := 4;
    ScenarioNoMatch : UINT := 5;
    ScenarioCaseSensitive : UINT := 6;
    ScenarioLongerFragment : UINT := 7;
    ScenarioEmptyInput : UINT := 8;
    ScenarioEmptyFragments : UINT := 9;
    ScenarioBothEmpty : UINT := 10;
    ScenarioIncompleteLastCandidate : UINT := 11;
    ScenarioWideCodeUnits : UINT := 12;
    ScenarioLastAtCapacity : UINT := 13;
    ScenarioWholeAtCapacity : UINT := 14;
    ScenarioInputOverCapacity : UINT := 15;
    ScenarioFragmentsOverCapacity : UINT := 16;
    LastScenario : UINT := ScenarioFragmentsOverCapacity;
END_VAR

SUPER^();

{region 'Documentation'}
(*!
<summary>Aggregates only outer checks, not intentionally failing subjects.</summary>
*)
{endregion}
METHOD PROTECTED AggregateResults
VAR_INPUT
    Aggregator : I_ResultAggregator; //! Borrowed result sink owned by the outer Test Case; add this test's checking Assertions without resetting or retaining the sink.
END_VAR
Aggregator.AddProvider(Provider := FResults);
Aggregator.AddProvider(Provider := FActivity);
Aggregator.AddProvider(Provider := FInputs);
Aggregator.AddProvider(Provider := FFindings);
END_METHOD

{region 'Documentation'}
(*!
<summary>Calls each inherited production subject once with caller-owned text storage.</summary>
*)
{endregion}
METHOD PRIVATE CallSubjects
FStartsWith(Enable := TRUE,
    State := E_State.Running,
    IN := FInput,
    Prefix := FPrefix);
FEndsWith(Enable := TRUE,
    State := E_State.Running,
    IN := FInput,
    Suffix := FSuffix);
FContains(Enable := TRUE,
    State := E_State.Running,
    IN := FInput,
    Fragment := FFragment);
FWideStartsWith(Enable := TRUE,
    State := E_State.Running,
    IN := FWideInput,
    Prefix := FWidePrefix);
FWideEndsWith(Enable := TRUE,
    State := E_State.Running,
    IN := FWideInput,
    Suffix := FWideSuffix);
FWideContains(Enable := TRUE,
    State := E_State.Running,
    IN := FWideInput,
    Fragment := FWideFragment);
END_METHOD

{region 'Documentation'}
(*!
<summary>Checks one subject finding in call order; expected outcomes come from the scenario.</summary>
*)
{endregion}
METHOD PRIVATE CheckFinding : BOOL //! TRUE when the required finding checks pass; calls requiring no finding also succeed.
VAR_INPUT
    Subject : I_Assertion; //! Assertion interface supplying the expected finding identity.
    ExpectedResult : E_Result; //! Independently authored result expected in the captured finding.
END_VAR
VAR_IN_OUT
    Index : UINT; //! One-based next finding index; advanced when this call checks a required finding.
END_VAR
CheckFinding := TRUE;
IF FEvaluateSubjects AND ((ExpectedResult = E_Result.Failed)
    OR (ExpectedResult = E_Result.Error)) THEN
    CheckFinding := (FEvents[Index].SequenceId = UINT_TO_UDINT(Index))
        AND (FEvents[Index].Name = Subject.Name)
        AND (FEvents[Index].OwnerScope = E_OwnerScope.Assertion)
        AND (FEvents[Index].EventType = E_EventType.Result)
        AND (FEvents[Index].State = E_State.Running)
        AND (FEvents[Index].Result = ExpectedResult)
        AND (FEvents[Index].Message <> '');
    Index := Index + 1;
END_IF;
END_METHOD

{region 'Documentation'}
(*!
<summary>Checks exact finding count and identities; at most one finding per subject.</summary>
*)
{endregion}
METHOD PRIVATE CheckFindings
VAR
    Index : UINT;
    Matches : BOOL;
END_VAR
Index := 1;
FFindingsMatch := TRUE;
Matches := CheckFinding(Subject := FStartsWith,
    ExpectedResult := FStartsWithExpectedResult,
    Index := Index);
FFindingsMatch := FFindingsMatch AND Matches;
Matches := CheckFinding(Subject := FEndsWith,
    ExpectedResult := FEndsWithExpectedResult,
    Index := Index);
FFindingsMatch := FFindingsMatch AND Matches;
Matches := CheckFinding(Subject := FContains,
    ExpectedResult := FContainsExpectedResult,
    Index := Index);
FFindingsMatch := FFindingsMatch AND Matches;
Matches := CheckFinding(Subject := FWideStartsWith,
    ExpectedResult := FWideStartsWithExpectedResult,
    Index := Index);
FFindingsMatch := FFindingsMatch AND Matches;
Matches := CheckFinding(Subject := FWideEndsWith,
    ExpectedResult := FWideEndsWithExpectedResult,
    Index := Index);
FFindingsMatch := FFindingsMatch AND Matches;
Matches := CheckFinding(Subject := FWideContains,
    ExpectedResult := FWideContainsExpectedResult,
    Index := Index);
FFindingsMatch := FFindingsMatch AND Matches;
FFindingsMatch := FFindingsMatch
    AND (FCaptureStatus.SequenceId = UINT_TO_UDINT(Index - 1))
    AND (FCaptureStatus.LostEventCount = 0);
END_METHOD

{region 'Documentation'}
(*!
<summary>Rejects incomplete subject, capture or outer Assertion setup.</summary>
*)
{endregion}
METHOD PROTECTED CheckInitialization : BOOL //! TRUE when the inherited initialization check and this concrete fixture check both accept the setup.
CheckInitialization := SUPER^.CheckInitialization();
IF NOT CheckInitialization THEN
    RETURN;
END_IF;

CheckInitialization := FSetupValid
    AND (Param_Assertions.AssertionStringLength >= 5)
    AND (Param_Assertions.AssertionWStringLength >= 5)
    AND (Param_Assertions.AssertionWStringLength < WideInputCapacity)
    AND FResults.IsInitialized
    AND FActivity.IsInitialized
    AND FInputs.IsInitialized
    AND FFindings.IsInitialized;
IF NOT CheckInitialization THEN
    EventPublisher.PublishEvent(Event := CreateFrameworkEvent(Name := Name,
        ResourceName := '',
        State := State,
        Severity := E_EventSeverity.Error,
        Message := 'Text selftest setup failed.'));
END_IF;
END_METHOD

{region 'Documentation'}
(*!
<summary>Checks literal evaluation results, or NotEvaluated on the reset call.</summary>
*)
{endregion}
METHOD PRIVATE CheckResults
IF FEvaluateSubjects THEN
    FResultsMatch := (FStartsWith.Result = FStartsWithExpectedResult)
        AND (FEndsWith.Result = FEndsWithExpectedResult)
        AND (FContains.Result = FContainsExpectedResult)
        AND (FWideStartsWith.Result = FWideStartsWithExpectedResult)
        AND (FWideEndsWith.Result = FWideEndsWithExpectedResult)
        AND (FWideContains.Result = FWideContainsExpectedResult);
ELSE
    FResultsMatch := (FStartsWith.Result = E_Result.NotEvaluated)
        AND (FEndsWith.Result = E_Result.NotEvaluated)
        AND (FContains.Result = E_Result.NotEvaluated)
        AND (FWideStartsWith.Result = E_Result.NotEvaluated)
        AND (FWideEndsWith.Result = E_Result.NotEvaluated)
        AND (FWideContains.Result = E_Result.NotEvaluated);
END_IF;
FActivityMatch := FStartsWith.Enabled
    AND (FStartsWith.ObservationActive = FEvaluateSubjects)
    AND (FStartsWith.EvaluationActive = FEvaluateSubjects)
    AND FEndsWith.Enabled
    AND (FEndsWith.ObservationActive = FEvaluateSubjects)
    AND (FEndsWith.EvaluationActive = FEvaluateSubjects)
    AND FContains.Enabled
    AND (FContains.ObservationActive = FEvaluateSubjects)
    AND (FContains.EvaluationActive = FEvaluateSubjects)
    AND FWideStartsWith.Enabled
    AND (FWideStartsWith.ObservationActive = FEvaluateSubjects)
    AND (FWideStartsWith.EvaluationActive = FEvaluateSubjects)
    AND FWideEndsWith.Enabled
    AND (FWideEndsWith.ObservationActive = FEvaluateSubjects)
    AND (FWideEndsWith.EvaluationActive = FEvaluateSubjects)
    AND FWideContains.Enabled
    AND (FWideContains.ObservationActive = FEvaluateSubjects)
    AND (FWideContains.EvaluationActive = FEvaluateSubjects);
END_METHOD

{region 'Documentation'}
(*!
<summary>Initializes outer checks and isolates intentional subject findings.</summary>
*)
{endregion}
METHOD PROTECTED Configure
VAR
    Initialized : BOOL;
END_VAR
FPreparationStateCount := 0;
FTestStateCount := 1;
FResults.Initialize(Parent := THIS^,
    AssertionName := 'Results');
FActivity.Initialize(Parent := THIS^,
    AssertionName := 'Activity');
FInputs.Initialize(Parent := THIS^,
    AssertionName := 'Inputs');
FFindings.Initialize(Parent := THIS^,
    AssertionName := 'Findings');
FSetupValid := FCapture.Initialize(Buffer := FEvents,
    FifoControl := FCaptureFifo,
    Status := FCaptureStatus);
FStartsWith.BindPublisher(Publisher := FCapture);
Initialized := FStartsWith.Initialize(Parent := THIS^,
    AssertionName := 'StartsWith');
FSetupValid := FSetupValid AND Initialized;
FEndsWith.BindPublisher(Publisher := FCapture);
Initialized := FEndsWith.Initialize(Parent := THIS^,
    AssertionName := 'EndsWith');
FSetupValid := FSetupValid AND Initialized;
FContains.BindPublisher(Publisher := FCapture);
Initialized := FContains.Initialize(Parent := THIS^,
    AssertionName := 'Contains');
FSetupValid := FSetupValid AND Initialized;
FWideStartsWith.BindPublisher(Publisher := FCapture);
Initialized := FWideStartsWith.Initialize(Parent := THIS^,
    AssertionName := 'WideStartsWith');
FSetupValid := FSetupValid AND Initialized;
FWideEndsWith.BindPublisher(Publisher := FCapture);
Initialized := FWideEndsWith.Initialize(Parent := THIS^,
    AssertionName := 'WideEndsWith');
FSetupValid := FSetupValid AND Initialized;
FWideContains.BindPublisher(Publisher := FCapture);
Initialized := FWideContains.Initialize(Parent := THIS^,
    AssertionName := 'WideContains');
FSetupValid := FSetupValid AND Initialized;
END_METHOD

{region 'Documentation'}
(*!
<summary>Completes abort; no asynchronous resource is owned.</summary>
*)
{endregion}
METHOD PROTECTED ProcessAbort
VAR_INPUT
    Enable : BOOL; //! Phase permission supplied by the owning Test Case; FALSE does not authorize progression, while observation may continue.
END_VAR
IF Enable THEN
    CompleteAbort();
END_IF;
END_METHOD

{region 'Documentation'}
(*!
<summary>Latches this call's checks before progression is permitted.</summary>
*)
{endregion}
METHOD PROTECTED ProcessAssertions
VAR_INPUT
    Enable : BOOL; //! Phase permission supplied by the owning Test Case; FALSE does not authorize progression, while observation may continue.
END_VAR
VAR
    Check : BOOL;
END_VAR
Check := Enable AND FObservationReady;
FResults(Enable := Check,
    State := State,
    IN := FResultsMatch);
FActivity(Enable := Check,
    State := State,
    IN := FActivityMatch);
FInputs(Enable := Check,
    State := State,
    IN := FInputsMatch);
FFindings(Enable := Check,
    State := State,
    IN := FFindingsMatch);
IF Check THEN
    FChecked := TRUE;
END_IF;
END_METHOD

{region 'Documentation'}
(*!
<summary>No Preparation phase is needed.</summary>
*)
{endregion}
METHOD PROTECTED ProcessPreparations
VAR_INPUT
    // SA0033: Required hook; this test has no Preparation phase.
    {attribute 'analysis' := '-33'}
    Enable : BOOL; //! Phase permission supplied by the owning Test Case; FALSE does not authorize progression, while observation may continue.
END_VAR
END_METHOD

{region 'Documentation'}
(*!
<summary>Restarts the scenario sequence and outer checks.</summary>
*)
{endregion}
METHOD PROTECTED ProcessReset
FScenario := ScenarioMatching;
FChecked := FALSE;
FEvaluateSubjects := FALSE;
FObservationReady := FALSE;
FFirstFailedScenario := 0;
FFailedDuringEvaluation := FALSE;
FCapture.Reset();
ResetSubjects();
FResults.Reset();
FActivity.Reset();
FInputs.Reset();
FFindings.Reset();
CompleteReset();
END_METHOD

{region 'Documentation'}
(*!
<summary>Resets then evaluates each scenario on separate cycles before advancing.</summary>
*)
{endregion}
METHOD PROTECTED ProcessTests
VAR_INPUT
    Enable : BOOL; //! Phase permission supplied by the owning Test Case; FALSE does not authorize progression, while observation may continue.
END_VAR
IF NOT Enable THEN
    RETURN;
END_IF;

IF FChecked THEN
    FChecked := FALSE;
    FObservationReady := FALSE;
    IF FEvaluateSubjects THEN
        IF FScenario = LastScenario THEN
            CompleteTests();
            RETURN;
        END_IF;
        FScenario := FScenario + 1;
    END_IF;
    FEvaluateSubjects := NOT FEvaluateSubjects;
END_IF;

IF NOT SelectScenario() THEN
    RETURN;
END_IF;
FCapture.Reset();
IF NOT FEvaluateSubjects THEN
    ResetSubjects();
END_IF;
FInputBefore := FInput;
FWideInputBefore := FWideInput;
FPrefixBefore := FPrefix;
FWidePrefixBefore := FWidePrefix;
FSuffixBefore := FSuffix;
FWideSuffixBefore := FWideSuffix;
FFragmentBefore := FFragment;
FWideFragmentBefore := FWideFragment;
CallSubjects();
CheckResults();
FInputsMatch := (FInput = FInputBefore)
    AND (FWideInput = FWideInputBefore)
    AND (FPrefix = FPrefixBefore)
    AND (FWidePrefix = FWidePrefixBefore)
    AND (FSuffix = FSuffixBefore)
    AND (FWideSuffix = FWideSuffixBefore)
    AND (FFragment = FFragmentBefore)
    AND (FWideFragment = FWideFragmentBefore);
CheckFindings();
IF (FFirstFailedScenario = 0)
    AND NOT (FResultsMatch AND FActivityMatch AND FInputsMatch AND FFindingsMatch) THEN
    FFirstFailedScenario := FScenario;
    FFailedDuringEvaluation := FEvaluateSubjects;
END_IF;
FObservationReady := TRUE;
END_METHOD

{region 'Documentation'}
(*!
<summary>Queues reset; the next bound FB call consumes it without evaluating.</summary>
*)
{endregion}
METHOD PRIVATE ResetSubjects
FStartsWith.Reset();
FEndsWith.Reset();
FContains.Reset();
FWideStartsWith.Reset();
FWideEndsWith.Reset();
FWideContains.Reset();
END_METHOD

{region 'Documentation'}
(*!
<summary>Selects explicit text stimuli and expected results for one scenario.</summary>
*)
{endregion}
METHOD PRIVATE SelectScenario : BOOL //! TRUE after selecting a supported scenario and its literal expectations; FALSE reports an unknown scenario.
VAR
    Index : UINT;
END_VAR
SelectScenario := FALSE;
FInput := 'ABABA';
FWideInput := "ABABA";
FPrefix := 'AB';
FSuffix := 'BA';
FFragment := 'ABA';
FWidePrefix := "AB";
FWideSuffix := "BA";
FWideFragment := "ABA";
CASE FScenario OF
    ScenarioMatching:

        FStartsWithExpectedResult := E_Result.Passed;
        FEndsWithExpectedResult := E_Result.Passed;
        FContainsExpectedResult := E_Result.Passed;
        FWideStartsWithExpectedResult := E_Result.Passed;
        FWideEndsWithExpectedResult := E_Result.Passed;
        FWideContainsExpectedResult := E_Result.Passed;
    ScenarioWholeInput:
        FPrefix := 'ABABA';
        FWidePrefix := "ABABA";
        FSuffix := 'ABABA';
        FWideSuffix := "ABABA";
        FFragment := 'ABABA';
        FWideFragment := "ABABA";
        FStartsWithExpectedResult := E_Result.Passed;
        FEndsWithExpectedResult := E_Result.Passed;
        FContainsExpectedResult := E_Result.Passed;
        FWideStartsWithExpectedResult := E_Result.Passed;
        FWideEndsWithExpectedResult := E_Result.Passed;
        FWideContainsExpectedResult := E_Result.Passed;
    ScenarioFirstPosition:
        FInput := 'ABAXY';
        FWideInput := "ABAXY";
        FPrefix := 'ABA';
        FWidePrefix := "ABA";
        FSuffix := 'ABA';
        FWideSuffix := "ABA";
        FFragment := 'ABA';
        FWideFragment := "ABA";
        FStartsWithExpectedResult := E_Result.Passed;
        FEndsWithExpectedResult := E_Result.Failed;
        FContainsExpectedResult := E_Result.Passed;
        FWideStartsWithExpectedResult := E_Result.Passed;
        FWideEndsWithExpectedResult := E_Result.Failed;
        FWideContainsExpectedResult := E_Result.Passed;
    ScenarioLastPosition:
        FInput := 'XYABA';
        FWideInput := "XYABA";
        FPrefix := 'ABA';
        FWidePrefix := "ABA";
        FSuffix := 'ABA';
        FWideSuffix := "ABA";
        FFragment := 'ABA';
        FWideFragment := "ABA";
        FStartsWithExpectedResult := E_Result.Failed;
        FEndsWithExpectedResult := E_Result.Passed;
        FContainsExpectedResult := E_Result.Passed;
        FWideStartsWithExpectedResult := E_Result.Failed;
        FWideEndsWithExpectedResult := E_Result.Passed;
        FWideContainsExpectedResult := E_Result.Passed;
    ScenarioNoMatch:
        FPrefix := 'Z';
        FWidePrefix := "Z";
        FSuffix := 'Z';
        FWideSuffix := "Z";
        FFragment := 'Z';
        FWideFragment := "Z";
        FStartsWithExpectedResult := E_Result.Failed;
        FEndsWithExpectedResult := E_Result.Failed;
        FContainsExpectedResult := E_Result.Failed;
        FWideStartsWithExpectedResult := E_Result.Failed;
        FWideEndsWithExpectedResult := E_Result.Failed;
        FWideContainsExpectedResult := E_Result.Failed;
    ScenarioCaseSensitive:
        FPrefix := 'aba';
        FWidePrefix := "aba";
        FSuffix := 'aba';
        FWideSuffix := "aba";
        FFragment := 'aba';
        FWideFragment := "aba";
        FStartsWithExpectedResult := E_Result.Failed;
        FEndsWithExpectedResult := E_Result.Failed;
        FContainsExpectedResult := E_Result.Failed;
        FWideStartsWithExpectedResult := E_Result.Failed;
        FWideEndsWithExpectedResult := E_Result.Failed;
        FWideContainsExpectedResult := E_Result.Failed;
    ScenarioLongerFragment:
        FPrefix := 'ABABAX';
        FWidePrefix := "ABABAX";
        FSuffix := 'ABABAX';
        FWideSuffix := "ABABAX";
        FFragment := 'ABABAX';
        FWideFragment := "ABABAX";
        FStartsWithExpectedResult := E_Result.Failed;
        FEndsWithExpectedResult := E_Result.Failed;
        FContainsExpectedResult := E_Result.Failed;
        FWideStartsWithExpectedResult := E_Result.Failed;
        FWideEndsWithExpectedResult := E_Result.Failed;
        FWideContainsExpectedResult := E_Result.Failed;
    ScenarioEmptyInput:
        FInput := '';
        FWideInput := "";
        FStartsWithExpectedResult := E_Result.Failed;
        FEndsWithExpectedResult := E_Result.Failed;
        FContainsExpectedResult := E_Result.Failed;
        FWideStartsWithExpectedResult := E_Result.Failed;
        FWideEndsWithExpectedResult := E_Result.Failed;
        FWideContainsExpectedResult := E_Result.Failed;
    ScenarioEmptyFragments:
        FPrefix := '';
        FWidePrefix := "";
        FSuffix := '';
        FWideSuffix := "";
        FFragment := '';
        FWideFragment := "";
        FStartsWithExpectedResult := E_Result.Error;
        FEndsWithExpectedResult := E_Result.Error;
        FContainsExpectedResult := E_Result.Error;
        FWideStartsWithExpectedResult := E_Result.Error;
        FWideEndsWithExpectedResult := E_Result.Error;
        FWideContainsExpectedResult := E_Result.Error;
    ScenarioBothEmpty:
        FInput := '';
        FWideInput := "";
        FPrefix := '';
        FWidePrefix := "";
        FSuffix := '';
        FWideSuffix := "";
        FFragment := '';
        FWideFragment := "";
        FStartsWithExpectedResult := E_Result.Error;
        FEndsWithExpectedResult := E_Result.Error;
        FContainsExpectedResult := E_Result.Error;
        FWideStartsWithExpectedResult := E_Result.Error;
        FWideEndsWithExpectedResult := E_Result.Error;
        FWideContainsExpectedResult := E_Result.Error;
    ScenarioIncompleteLastCandidate:
        FInput := 'XYAB';
        FWideInput := "XYAB";
        FPrefix := 'ABC';
        FWidePrefix := "ABC";
        FSuffix := 'ABC';
        FWideSuffix := "ABC";
        FFragment := 'ABC';
        FWideFragment := "ABC";
        FStartsWithExpectedResult := E_Result.Failed;
        FEndsWithExpectedResult := E_Result.Failed;
        FContainsExpectedResult := E_Result.Failed;
        FWideStartsWithExpectedResult := E_Result.Failed;
        FWideEndsWithExpectedResult := E_Result.Failed;
        FWideContainsExpectedResult := E_Result.Failed;
    ScenarioWideCodeUnits:
        FWideInput := "ABC";
        FWideInput[0] := WORD#16#0100;
        FWideInput[1] := WORD#16#0141;
        FWidePrefix := "A";
        FWidePrefix[0] := WORD#16#0100;
        FWideSuffix := "AC";
        FWideSuffix[0] := WORD#16#0141;
        FWideFragment := "A";
        FWideFragment[0] := WORD#16#0241;
        FStartsWithExpectedResult := E_Result.Passed;
        FEndsWithExpectedResult := E_Result.Passed;
        FContainsExpectedResult := E_Result.Passed;
        FWideStartsWithExpectedResult := E_Result.Passed;
        FWideEndsWithExpectedResult := E_Result.Passed;
        FWideContainsExpectedResult := E_Result.Failed;
    ScenarioLastAtCapacity:
        FOR Index := 0 TO Param_Assertions.AssertionStringLength - 1 DO
            // SA0175: Bounded byte writes construct exact input/terminator boundaries; no UTF-8 decoding.
            {analysis -175}
            FInput[Index] := BYTE#16#41;
            {analysis +175}
        END_FOR;
        // SA0175: Bounded byte writes construct exact input/terminator boundaries; no UTF-8 decoding.
        {analysis -175}
        FInput[Param_Assertions.AssertionStringLength - 1] := BYTE#16#5A;
        FInput[Param_Assertions.AssertionStringLength] := 0;
        {analysis +175}
        FOR Index := 0 TO Param_Assertions.AssertionWStringLength - 1 DO
            FWideInput[Index] := WORD#16#0141;
        END_FOR;
        FWideInput[Param_Assertions.AssertionWStringLength - 1] := WORD#16#0100;
        FWideInput[Param_Assertions.AssertionWStringLength] := 0;
        FPrefix := 'A';
        FSuffix := 'Z';
        FFragment := 'AZ';
        FWidePrefix := "A";
        FWidePrefix[0] := WORD#16#0141;
        FWideSuffix := "Z";
        FWideSuffix[0] := WORD#16#0100;
        FWideFragment := "AZ";
        FWideFragment[0] := WORD#16#0141;
        FWideFragment[1] := WORD#16#0100;
        FStartsWithExpectedResult := E_Result.Passed;
        FEndsWithExpectedResult := E_Result.Passed;
        FContainsExpectedResult := E_Result.Passed;
        FWideStartsWithExpectedResult := E_Result.Passed;
        FWideEndsWithExpectedResult := E_Result.Passed;
        FWideContainsExpectedResult := E_Result.Passed;
    ScenarioWholeAtCapacity:
        FOR Index := 0 TO Param_Assertions.AssertionStringLength - 1 DO
            // SA0175: Bounded byte writes construct exact input/terminator boundaries; no UTF-8 decoding.
            {analysis -175}
            FInput[Index] := BYTE#16#41;
            {analysis +175}
        END_FOR;
        // SA0175: Bounded byte writes construct exact input/terminator boundaries; no UTF-8 decoding.
        {analysis -175}
        FInput[Param_Assertions.AssertionStringLength - 1] := BYTE#16#5A;
        FInput[Param_Assertions.AssertionStringLength] := 0;
        {analysis +175}
        FOR Index := 0 TO Param_Assertions.AssertionWStringLength - 1 DO
            FWideInput[Index] := WORD#16#0141;
        END_FOR;
        FWideInput[Param_Assertions.AssertionWStringLength - 1] := WORD#16#0100;
        FWideInput[Param_Assertions.AssertionWStringLength] := 0;
        FPrefix := 'A';
        FSuffix := 'Z';
        FFragment := 'AZ';
        FWidePrefix := "A";
        FWidePrefix[0] := WORD#16#0141;
        FWideSuffix := "Z";
        FWideSuffix[0] := WORD#16#0100;
        FWideFragment := "AZ";
        FWideFragment[0] := WORD#16#0141;
        FWideFragment[1] := WORD#16#0100;
        FPrefix := FInput;
        FSuffix := FInput;
        FFragment := FInput;
        FWidePrefix := FWideInput;
        FWideSuffix := FWideInput;
        FWideFragment := FWideInput;
        FStartsWithExpectedResult := E_Result.Passed;
        FEndsWithExpectedResult := E_Result.Passed;
        FContainsExpectedResult := E_Result.Passed;
        FWideStartsWithExpectedResult := E_Result.Passed;
        FWideEndsWithExpectedResult := E_Result.Passed;
        FWideContainsExpectedResult := E_Result.Passed;
    ScenarioInputOverCapacity:
        FOR Index := 0 TO Param_Assertions.AssertionStringLength - 1 DO
            // SA0175: Bounded byte writes construct exact input/terminator boundaries; no UTF-8 decoding.
            {analysis -175}
            FInput[Index] := BYTE#16#41;
            {analysis +175}
        END_FOR;
        // SA0175: Bounded byte writes construct exact input/terminator boundaries; no UTF-8 decoding.
        {analysis -175}
        FInput[Param_Assertions.AssertionStringLength - 1] := BYTE#16#5A;
        FInput[Param_Assertions.AssertionStringLength] := 0;
        {analysis +175}
        FOR Index := 0 TO Param_Assertions.AssertionWStringLength - 1 DO
            FWideInput[Index] := WORD#16#0141;
        END_FOR;
        FWideInput[Param_Assertions.AssertionWStringLength - 1] := WORD#16#0100;
        FWideInput[Param_Assertions.AssertionWStringLength] := 0;
        FPrefix := 'A';
        FSuffix := 'Z';
        FFragment := 'AZ';
        FWidePrefix := "A";
        FWidePrefix[0] := WORD#16#0141;
        FWideSuffix := "Z";
        FWideSuffix[0] := WORD#16#0100;
        FWideFragment := "AZ";
        FWideFragment[0] := WORD#16#0141;
        FWideFragment[1] := WORD#16#0100;
        // SA0175: Bounded byte writes construct exact input/terminator boundaries; no UTF-8 decoding.
        {analysis -175}
        FInput[Param_Assertions.AssertionStringLength] := BYTE#16#41;
        FInput[Param_Assertions.AssertionStringLength + 1] := 0;
        {analysis +175}
        FWideInput[Param_Assertions.AssertionWStringLength] := WORD#16#0141;
        FWideInput[Param_Assertions.AssertionWStringLength + 1] := 0;
        FStartsWithExpectedResult := E_Result.Error;
        FEndsWithExpectedResult := E_Result.Error;
        FContainsExpectedResult := E_Result.Error;
        FWideStartsWithExpectedResult := E_Result.Error;
        FWideEndsWithExpectedResult := E_Result.Error;
        FWideContainsExpectedResult := E_Result.Error;
    ScenarioFragmentsOverCapacity:
        FOR Index := 0 TO Param_Assertions.AssertionStringLength - 1 DO
            // SA0175: Bounded byte writes construct exact input/terminator boundaries; no UTF-8 decoding.
            {analysis -175}
            FInput[Index] := BYTE#16#41;
            {analysis +175}
        END_FOR;
        // SA0175: Bounded byte writes construct exact input/terminator boundaries; no UTF-8 decoding.
        {analysis -175}
        FInput[Param_Assertions.AssertionStringLength - 1] := BYTE#16#5A;
        FInput[Param_Assertions.AssertionStringLength] := 0;
        {analysis +175}
        FOR Index := 0 TO Param_Assertions.AssertionWStringLength - 1 DO
            FWideInput[Index] := WORD#16#0141;
        END_FOR;
        FWideInput[Param_Assertions.AssertionWStringLength - 1] := WORD#16#0100;
        FWideInput[Param_Assertions.AssertionWStringLength] := 0;
        FPrefix := 'A';
        FSuffix := 'Z';
        FFragment := 'AZ';
        FWidePrefix := "A";
        FWidePrefix[0] := WORD#16#0141;
        FWideSuffix := "Z";
        FWideSuffix[0] := WORD#16#0100;
        FWideFragment := "AZ";
        FWideFragment[0] := WORD#16#0141;
        FWideFragment[1] := WORD#16#0100;
        // SA0175: Bounded byte writes construct exact input/terminator boundaries; no UTF-8 decoding.
        {analysis -175}
        FInput[Param_Assertions.AssertionStringLength] := BYTE#16#41;
        FInput[Param_Assertions.AssertionStringLength + 1] := 0;
        {analysis +175}
        FWideInput[Param_Assertions.AssertionWStringLength] := WORD#16#0141;
        FWideInput[Param_Assertions.AssertionWStringLength + 1] := 0;
        FPrefix := FInput;
        FSuffix := FInput;
        FFragment := FInput;
        FWidePrefix := FWideInput;
        FWideSuffix := FWideInput;
        FWideFragment := FWideInput;
        FInput := 'A';
        FWideInput := "A";
        FStartsWithExpectedResult := E_Result.Error;
        FEndsWithExpectedResult := E_Result.Error;
        FContainsExpectedResult := E_Result.Error;
        FWideStartsWithExpectedResult := E_Result.Error;
        FWideEndsWithExpectedResult := E_Result.Error;
        FWideContainsExpectedResult := E_Result.Error;
ELSE
    Error(Message := 'Unknown text scenario.');
    RETURN;
END_CASE;
SelectScenario := TRUE;
END_METHOD

END_FUNCTION_BLOCK

// ---- SelfTests/TestCases/TestSuite_AssertionText/Test_AssertionTextDiagnostics.TcPOU
{region 'Documentation'}
(*!
<summary>Checks complete Failed-event messages, quoted previews and character code fallbacks.</summary>
<description>
Text and character Assertions publish into a local capture. Expected messages
are literal independent examples, not outputs from the formatter under test.
Preview boundaries use the contract limit of 40 output bytes; a difference
beyond the preview still fails even when both rendered previews are identical.
Independent scenarios occupy two calls: bound Reset, then evaluation.
ProcessAssertions checks each call before ProcessTests advances. Literal expected
results belong to SelectScenario, not to a copy of the production comparison.
The local capture is cleared before each call and checked in subject-call order.
FirstFailedScenario and FailedDuringEvaluation retain the first mismatch.
Continuation scenarios explicitly retain the prior subject state. The Test Case
owns all input storage; no invalid or dangling references are constructed.
</description>
*)
{endregion}
FUNCTION_BLOCK Test_AssertionTextDiagnostics EXTENDS TestCaseBase
VAR
    FText : AssertEqual_String;
    FTextExpectedResult : E_Result;
    FWideText : AssertEqual_WString;
    FWideTextExpectedResult : E_Result;
    FCharacter : AssertEqual_Char;
    FCharacterExpectedResult : E_Result;
    FWideCharacter : AssertEqual_WChar;
    FWideCharacterExpectedResult : E_Result;
    FInput : STRING(Param_Assertions.AssertionStringLength);
    FInputBefore : STRING(Param_Assertions.AssertionStringLength);
    FExpected : STRING(Param_Assertions.AssertionStringLength);
    FExpectedBefore : STRING(Param_Assertions.AssertionStringLength);
    FWideInput : WSTRING(Param_Assertions.AssertionWStringLength);
    FWideInputBefore : WSTRING(Param_Assertions.AssertionWStringLength);
    FWideExpected : WSTRING(Param_Assertions.AssertionWStringLength);
    FWideExpectedBefore : WSTRING(Param_Assertions.AssertionWStringLength);
    FChar : BYTE;
    FCharBefore : BYTE;
    FExpectedChar : BYTE;
    FExpectedCharBefore : BYTE;
    FWideChar : WORD;
    FWideCharBefore : WORD;
    FExpectedWideChar : WORD;
    FExpectedWideCharBefore : WORD;
    FExpectedMessage1 : STRING(GVL_Constants.MessageLength);
    FExpectedMessage2 : STRING(GVL_Constants.MessageLength);
    FExpectedMessage3 : STRING(GVL_Constants.MessageLength);
    FExpectedMessage4 : STRING(GVL_Constants.MessageLength);
    FSubjectEnable : BOOL;
    FContinueScenario : BOOL;
    FTextExpectedFinding : BOOL;
    FWideTextExpectedFinding : BOOL;
    FCharacterExpectedFinding : BOOL;
    FWideCharacterExpectedFinding : BOOL;
    FCapture : EventBuffer;
    FEvents : ARRAY[1..CaptureLength] OF ST_Event;
    FCaptureFifo : ST_FifoStatus;
    FCaptureStatus : ST_EventBufferStatus;
    FSetupValid : BOOL;
    FScenario : UINT;
    FChecked : BOOL;
    FEvaluateSubjects : BOOL;
    FObservationReady : BOOL;
    FFirstFailedScenario : UINT;
    FFailedDuringEvaluation : BOOL;
    FResultsMatch : BOOL;
    FResults : AssertTrue;
    FActivityMatch : BOOL;
    FActivity : AssertTrue;
    FInputsMatch : BOOL;
    FInputs : AssertTrue;
    FFindingsMatch : BOOL;
    FPreviewRenderingMatch : BOOL;
    FFindings : AssertTrue;
END_VAR
VAR CONSTANT
    CaptureLength : UINT := 8;
    ScenarioShortQuoted : UINT := 1;
    ScenarioPreview38 : UINT := 2;
    ScenarioPreview39 : UINT := 3;
    ScenarioDifferenceBeyondPreview : UINT := 4;
    ScenarioAtCapacity : UINT := 5;
    ScenarioCodeFallback : UINT := 6;
    ScenarioReplacement : UINT := 7;
    LastScenario : UINT := ScenarioReplacement;
END_VAR

SUPER^();

{region 'Documentation'}
(*!
<summary>Aggregates only outer checks, not intentionally failing subjects.</summary>
*)
{endregion}
METHOD PROTECTED AggregateResults
VAR_INPUT
    Aggregator : I_ResultAggregator; //! Borrowed result sink owned by the outer Test Case; add this test's checking Assertions without resetting or retaining the sink.
END_VAR
Aggregator.AddProvider(Provider := FResults);
Aggregator.AddProvider(Provider := FActivity);
Aggregator.AddProvider(Provider := FInputs);
Aggregator.AddProvider(Provider := FFindings);
END_METHOD

{region 'Documentation'}
(*!
<summary>Calls each inherited production subject once with caller-owned input storage.</summary>
*)
{endregion}
METHOD PRIVATE CallSubjects
FText(Enable := FSubjectEnable,
    State := E_State.Running,
    IN := FInput,
    Expected := FExpected);
FWideText(Enable := FSubjectEnable,
    State := E_State.Running,
    IN := FWideInput,
    Expected := FWideExpected);
FCharacter(Enable := FSubjectEnable,
    State := E_State.Running,
    IN := FChar,
    Expected := FExpectedChar);
FWideCharacter(Enable := FSubjectEnable,
    State := E_State.Running,
    IN := FWideChar,
    Expected := FExpectedWideChar);
END_METHOD

{region 'Documentation'}
(*!
<summary>Checks one subject finding in call order; expected outcomes come from the scenario.</summary>
*)
{endregion}
METHOD PRIVATE CheckFinding : BOOL //! TRUE when the required finding checks pass; calls requiring no finding also succeed.
VAR_INPUT
    Subject : I_Assertion; //! Assertion interface supplying the expected finding identity.
    ExpectedResult : E_Result; //! Independently authored result expected in the captured finding.
    ExpectedFinding : BOOL; //! TRUE when this scenario requires a finding during active evaluation.
END_VAR
VAR_IN_OUT
    Index : UINT; //! One-based next finding index; advanced when this call checks a required finding.
END_VAR
CheckFinding := TRUE;
IF FEvaluateSubjects AND ExpectedFinding THEN
    CheckFinding := (FEvents[Index].SequenceId = UINT_TO_UDINT(Index))
        AND (FEvents[Index].Name = Subject.Name)
        AND (FEvents[Index].OwnerScope = E_OwnerScope.Assertion)
        AND (FEvents[Index].EventType = E_EventType.Result)
        AND (FEvents[Index].State = E_State.Running)
        AND (FEvents[Index].Result = ExpectedResult)
        AND (FEvents[Index].Message <> '');
    Index := Index + 1;
END_IF;
END_METHOD

{region 'Documentation'}
(*!
<summary>Checks exact finding count and identities; at most one finding per subject.</summary>
*)
{endregion}
METHOD PRIVATE CheckFindings
VAR
    Index : UINT;
    Matches : BOOL;
END_VAR
Index := 1;
FFindingsMatch := TRUE;
Matches := CheckFinding(Subject := FText,
    ExpectedResult := FTextExpectedResult,
    ExpectedFinding := FTextExpectedFinding,
    Index := Index);
FFindingsMatch := FFindingsMatch AND Matches;
Matches := CheckFinding(Subject := FWideText,
    ExpectedResult := FWideTextExpectedResult,
    ExpectedFinding := FWideTextExpectedFinding,
    Index := Index);
FFindingsMatch := FFindingsMatch AND Matches;
Matches := CheckFinding(Subject := FCharacter,
    ExpectedResult := FCharacterExpectedResult,
    ExpectedFinding := FCharacterExpectedFinding,
    Index := Index);
FFindingsMatch := FFindingsMatch AND Matches;
Matches := CheckFinding(Subject := FWideCharacter,
    ExpectedResult := FWideCharacterExpectedResult,
    ExpectedFinding := FWideCharacterExpectedFinding,
    Index := Index);
FFindingsMatch := FFindingsMatch AND Matches;
FFindingsMatch := FFindingsMatch
    AND (FCaptureStatus.SequenceId = UINT_TO_UDINT(Index - 1))
    AND (FCaptureStatus.LostEventCount = 0);
IF FEvaluateSubjects THEN
    FFindingsMatch := FFindingsMatch
        AND (FEvents[1].Message = FExpectedMessage1)
        AND (LEN(FEvents[1].Message) <= GVL_Constants.MessageLength)
        AND (FEvents[2].Message = FExpectedMessage2)
        AND (LEN(FEvents[2].Message) <= GVL_Constants.MessageLength)
        AND (FEvents[3].Message = FExpectedMessage3)
        AND (LEN(FEvents[3].Message) <= GVL_Constants.MessageLength)
        AND (FEvents[4].Message = FExpectedMessage4)
        AND (LEN(FEvents[4].Message) <= GVL_Constants.MessageLength);
END_IF;
END_METHOD

{region 'Documentation'}
(*!
<summary>Rejects incomplete subject, capture or outer Assertion setup.</summary>
*)
{endregion}
METHOD PROTECTED CheckInitialization : BOOL //! TRUE when the inherited initialization check and this concrete fixture check both accept the setup.
CheckInitialization := SUPER^.CheckInitialization();
IF NOT CheckInitialization THEN
    RETURN;
END_IF;

CheckInitialization := FSetupValid
    AND (GVL_Constants.AssertionValueLength = 40)
    AND (Param_Assertions.AssertionStringLength >= 40)
    AND (Param_Assertions.AssertionWStringLength >= 40)
    AND FResults.IsInitialized
    AND FActivity.IsInitialized
    AND FInputs.IsInitialized
    AND FFindings.IsInitialized;
IF NOT CheckInitialization THEN
    EventPublisher.PublishEvent(Event := CreateFrameworkEvent(Name := Name,
        ResourceName := '',
        State := State,
        Severity := E_EventSeverity.Error,
        Message := 'Text selftest setup failed.'));
END_IF;
END_METHOD

{region 'Documentation'}
(*!
<summary>Checks literal replacement, terminator, array-zero and preview-boundary examples.</summary>
<description>
Exercises all four production preview functions directly, including negative array
bounds and unchanged input storage. Expected bytes are authored independently.
The existing event scenarios separately check comparison results and publication.
</description>
*)
{endregion}
METHOD PRIVATE CheckPreviewRendering : BOOL //! TRUE when every literal preview and input-preservation check succeeds.
VAR
    Matches : BOOL;
    Text : STRING(40);
    WideText : WSTRING(40);
    Bytes : ARRAY[-2..37] OF BYTE;
    Words : ARRAY[-2..37] OF WORD;
    Index : DINT;
END_VAR
Matches := TRUE;
// SA0175: Deliberate byte fixtures and literal expected transport bytes, not UTF-8 text.
{analysis -175}
Text := '$01$1F$7F$80$D7$FF';
WideText := "$0001$001F$007F$0080$0100$20AC";
Matches := Matches AND (CreateAssertionTextValue_String(Value := Text) = '$'$D7$D7$D7$D7$D7$D7$'');
Matches := Matches AND (CreateAssertionTextValue_WString(Value := WideText) = '$'$D7$D7$D7$D7$D7$D7$'');
Matches := Matches AND (Text = '$01$1F$7F$80$D7$FF');
Matches := Matches AND (WideText = "$0001$001F$007F$0080$0100$20AC");

Text := ' ~$'\';
WideText := " ~$'\";
Matches := Matches AND (CreateAssertionTextValue_String(Value := Text) = '$' ~$'\$'');
Matches := Matches AND (CreateAssertionTextValue_WString(Value := WideText) = '$' ~$'\$'');
Matches := Matches AND (CreateAssertionTextValue_String(Value := '') = '$'$'');
Matches := Matches AND (CreateAssertionTextValue_WString(Value := "") = '$'$'');
Text := 'A$00B';
WideText := "A$0000B";
Matches := Matches AND (CreateAssertionTextValue_String(Value := Text) = '$'A$'');
Matches := Matches AND (CreateAssertionTextValue_WString(Value := WideText) = '$'A$'');

FOR Index := -2 TO 37 DO
    Bytes[Index] := BYTE#16#41;
    Words[Index] := WORD#16#0041;
END_FOR;
Matches := Matches AND (CreateAssertionTextValue_ByteArray(Value := Bytes, StartIndex := -2, Length := 38) = '$'AAAAAAAAAAAAAAAAAAAAAAAAAAAAAAAAAAAAAA$'');
Matches := Matches AND (CreateAssertionTextValue_WordArray(Value := Words, StartIndex := -2, Length := 38) = '$'AAAAAAAAAAAAAAAAAAAAAAAAAAAAAAAAAAAAAA$'');
Matches := Matches AND (CreateAssertionTextValue_ByteArray(Value := Bytes, StartIndex := -2, Length := 39) = '$'AAAAAAAAAAAAAAAAAAAAAAAAAAAAAAAAAAA...$'');
Matches := Matches AND (CreateAssertionTextValue_WordArray(Value := Words, StartIndex := -2, Length := 39) = '$'AAAAAAAAAAAAAAAAAAAAAAAAAAAAAAAAAAA...$'');
Text := 'AAAAAAAAAAAAAAAAAAAAAAAAAAAAAAAAAAAAA$FF';
WideText := "AAAAAAAAAAAAAAAAAAAAAAAAAAAAAAAAAAAAA$0100";
Matches := Matches AND (CreateAssertionTextValue_String(Value := Text) = '$'AAAAAAAAAAAAAAAAAAAAAAAAAAAAAAAAAAAAA$D7$'');
Matches := Matches AND (CreateAssertionTextValue_WString(Value := WideText) = '$'AAAAAAAAAAAAAAAAAAAAAAAAAAAAAAAAAAAAA$D7$'');
Text := 'AAAAAAAAAAAAAAAAAAAAAAAAAAAAAAAAAA$FFAAAA';
WideText := "AAAAAAAAAAAAAAAAAAAAAAAAAAAAAAAAAA$20ACAAAA";
Matches := Matches AND (CreateAssertionTextValue_String(Value := Text) = '$'AAAAAAAAAAAAAAAAAAAAAAAAAAAAAAAAAA$D7...$'');
Matches := Matches AND (CreateAssertionTextValue_WString(Value := WideText) = '$'AAAAAAAAAAAAAAAAAAAAAAAAAAAAAAAAAA$D7...$'');

Bytes[-2] := BYTE#16#20;
Bytes[-1] := 0;
Bytes[0] := BYTE#16#7E;
Bytes[1] := BYTE#16#E4;
Bytes[2] := BYTE#16#FF;
Bytes[3] := BYTE#16#1F;
Words[-2] := WORD#16#0020;
Words[-1] := 0;
Words[0] := WORD#16#007E;
Words[1] := WORD#16#0100;
Words[2] := WORD#16#20AC;
Words[3] := WORD#16#001F;
Matches := Matches AND (CreateAssertionTextValue_ByteArray(Value := Bytes, StartIndex := -2, Length := 6) = '$' $D7~$D7$D7$D7$'');
Matches := Matches AND (CreateAssertionTextValue_WordArray(Value := Words, StartIndex := -2, Length := 6) = '$' $D7~$D7$D7$D7$'');
Matches := Matches AND (Bytes[-2] = 16#20) AND (Bytes[-1] = 0) AND (Bytes[0] = 16#7E)
    AND (Bytes[1] = 16#E4) AND (Bytes[2] = 16#FF) AND (Bytes[3] = 16#1F);
Matches := Matches AND (Words[-2] = 16#20) AND (Words[-1] = 0) AND (Words[0] = 16#7E)
    AND (Words[1] = 16#0100) AND (Words[2] = 16#20AC) AND (Words[3] = 16#1F);
FOR Index := 4 TO 37 DO
    Matches := Matches AND (Bytes[Index] = 16#41) AND (Words[Index] = 16#41);
END_FOR;
Matches := Matches AND (CreateAssertionTextValue_ByteArray(Value := Bytes, StartIndex := -3, Length := 1) = '$'$'');
Matches := Matches AND (CreateAssertionTextValue_WordArray(Value := Words, StartIndex := 37, Length := 2) = '$'$'');
Matches := Matches AND (CreateAssertionTextValue_ByteArray(Value := Bytes, StartIndex := -2, Length := 0) = '$'$'');
Matches := Matches AND (CreateAssertionTextValue_WordArray(Value := Words, StartIndex := -2, Length := 0) = '$'$'');
{analysis +175}
Matches := Matches AND (CreateAssertionTextValue_Char(Value := 16#20) = '$' $' (16#20)');
Matches := Matches AND (CreateAssertionTextValue_Char(Value := 16#7E) = '$'~$' (16#7E)');
Matches := Matches AND (CreateAssertionTextValue_WChar(Value := 16#20) = '$' $' (16#0020)');
Matches := Matches AND (CreateAssertionTextValue_WChar(Value := 16#7E) = '$'~$' (16#007E)');
Matches := Matches AND (CreateAssertionTextValue_Char(Value := 16#FF) = '16#FF');
Matches := Matches AND (CreateAssertionTextValue_WChar(Value := 16#FFFF) = '16#FFFF');
CheckPreviewRendering := Matches;
END_METHOD

{region 'Documentation'}
(*!
<summary>Checks literal evaluation results, or NotEvaluated on the reset call.</summary>
*)
{endregion}
METHOD PRIVATE CheckResults
IF FEvaluateSubjects THEN
    FResultsMatch := (FText.Result = FTextExpectedResult)
        AND (FWideText.Result = FWideTextExpectedResult)
        AND (FCharacter.Result = FCharacterExpectedResult)
        AND (FWideCharacter.Result = FWideCharacterExpectedResult);
ELSE
    FResultsMatch := (FText.Result = E_Result.NotEvaluated)
        AND (FWideText.Result = E_Result.NotEvaluated)
        AND (FCharacter.Result = E_Result.NotEvaluated)
        AND (FWideCharacter.Result = E_Result.NotEvaluated);
END_IF;
FActivityMatch := (FText.Enabled = FSubjectEnable)
    AND (FText.ObservationActive = (FEvaluateSubjects AND FSubjectEnable))
    AND (FText.EvaluationActive = (FEvaluateSubjects AND FSubjectEnable))
    AND (FWideText.Enabled = FSubjectEnable)
    AND (FWideText.ObservationActive = (FEvaluateSubjects AND FSubjectEnable))
    AND (FWideText.EvaluationActive = (FEvaluateSubjects AND FSubjectEnable))
    AND (FCharacter.Enabled = FSubjectEnable)
    AND (FCharacter.ObservationActive = (FEvaluateSubjects AND FSubjectEnable))
    AND (FCharacter.EvaluationActive = (FEvaluateSubjects AND FSubjectEnable))
    AND (FWideCharacter.Enabled = FSubjectEnable)
    AND (FWideCharacter.ObservationActive = (FEvaluateSubjects AND FSubjectEnable))
    AND (FWideCharacter.EvaluationActive = (FEvaluateSubjects AND FSubjectEnable));
END_METHOD

{region 'Documentation'}
(*!
<summary>Initializes outer checks and isolates intentional subject findings.</summary>
*)
{endregion}
METHOD PROTECTED Configure
VAR
    Initialized : BOOL;
END_VAR
FPreparationStateCount := 0;
FTestStateCount := 1;
FResults.Initialize(Parent := THIS^,
    AssertionName := 'Results');
FActivity.Initialize(Parent := THIS^,
    AssertionName := 'Activity');
FInputs.Initialize(Parent := THIS^,
    AssertionName := 'Inputs');
FFindings.Initialize(Parent := THIS^,
    AssertionName := 'Findings');
FSetupValid := FCapture.Initialize(Buffer := FEvents,
    FifoControl := FCaptureFifo,
    Status := FCaptureStatus);
FText.BindPublisher(Publisher := FCapture);
Initialized := FText.Initialize(Parent := THIS^,
    AssertionName := 'Text');
FSetupValid := FSetupValid AND Initialized;
FWideText.BindPublisher(Publisher := FCapture);
Initialized := FWideText.Initialize(Parent := THIS^,
    AssertionName := 'WideText');
FSetupValid := FSetupValid AND Initialized;
FCharacter.BindPublisher(Publisher := FCapture);
Initialized := FCharacter.Initialize(Parent := THIS^,
    AssertionName := 'Character');
FSetupValid := FSetupValid AND Initialized;
FWideCharacter.BindPublisher(Publisher := FCapture);
Initialized := FWideCharacter.Initialize(Parent := THIS^,
    AssertionName := 'WideCharacter');
FSetupValid := FSetupValid AND Initialized;
END_METHOD

{region 'Documentation'}
(*!
<summary>Completes abort; no asynchronous resource is owned.</summary>
*)
{endregion}
METHOD PROTECTED ProcessAbort
VAR_INPUT
    Enable : BOOL; //! Phase permission supplied by the owning Test Case; FALSE does not authorize progression, while observation may continue.
END_VAR
IF Enable THEN
    CompleteAbort();
END_IF;
END_METHOD

{region 'Documentation'}
(*!
<summary>Latches this call's checks before progression is permitted.</summary>
*)
{endregion}
METHOD PROTECTED ProcessAssertions
VAR_INPUT
    Enable : BOOL; //! Phase permission supplied by the owning Test Case; FALSE does not authorize progression, while observation may continue.
END_VAR
VAR
    Check : BOOL;
END_VAR
Check := Enable AND FObservationReady;
FResults(Enable := Check,
    State := State,
    IN := FResultsMatch);
FActivity(Enable := Check,
    State := State,
    IN := FActivityMatch);
FInputs(Enable := Check,
    State := State,
    IN := FInputsMatch);
FFindings(Enable := Check,
    State := State,
    IN := FFindingsMatch);
IF Check THEN
    FChecked := TRUE;
END_IF;
END_METHOD

{region 'Documentation'}
(*!
<summary>No Preparation phase is needed.</summary>
*)
{endregion}
METHOD PROTECTED ProcessPreparations
VAR_INPUT
    // SA0033: Required hook; this test has no Preparation phase.
    {attribute 'analysis' := '-33'}
    Enable : BOOL; //! Phase permission supplied by the owning Test Case; FALSE does not authorize progression, while observation may continue.
END_VAR
END_METHOD

{region 'Documentation'}
(*!
<summary>Restarts the scenario sequence and outer checks.</summary>
*)
{endregion}
METHOD PROTECTED ProcessReset
FScenario := ScenarioShortQuoted;
FPreviewRenderingMatch := TRUE;
FChecked := FALSE;
FSubjectEnable := FALSE;
FContinueScenario := FALSE;
FEvaluateSubjects := FALSE;
FObservationReady := FALSE;
FFirstFailedScenario := 0;
FFailedDuringEvaluation := FALSE;
FCapture.Reset();
ResetSubjects();
FResults.Reset();
FActivity.Reset();
FInputs.Reset();
FFindings.Reset();
CompleteReset();
END_METHOD

{region 'Documentation'}
(*!
<summary>Consumes reset before each independent scenario; continuation retains subject state.</summary>
*)
{endregion}
METHOD PROTECTED ProcessTests
VAR_INPUT
    Enable : BOOL; //! Phase permission supplied by the owning Test Case; FALSE does not authorize progression, while observation may continue.
END_VAR
IF NOT Enable THEN
    RETURN;
END_IF;

IF FChecked THEN
    FChecked := FALSE;
    FObservationReady := FALSE;
    IF FEvaluateSubjects THEN
        IF FScenario = LastScenario THEN
            CompleteTests();
            RETURN;
        END_IF;
        FScenario := FScenario + 1;
    END_IF;
    FEvaluateSubjects := NOT FEvaluateSubjects;
END_IF;

IF NOT SelectScenario() THEN
    RETURN;
END_IF;
IF FContinueScenario THEN
    FEvaluateSubjects := TRUE;
END_IF;
FCapture.Reset();
IF NOT FEvaluateSubjects THEN
    ResetSubjects();
END_IF;
FInputBefore := FInput;
FExpectedBefore := FExpected;
FWideInputBefore := FWideInput;
FWideExpectedBefore := FWideExpected;
FCharBefore := FChar;
FExpectedCharBefore := FExpectedChar;
FWideCharBefore := FWideChar;
FExpectedWideCharBefore := FExpectedWideChar;
IF FScenario = ScenarioShortQuoted THEN
    FPreviewRenderingMatch := CheckPreviewRendering();
END_IF;
CallSubjects();
CheckResults();
FInputsMatch := (FInput = FInputBefore)
    AND (FExpected = FExpectedBefore)
    AND (FWideInput = FWideInputBefore)
    AND (FWideExpected = FWideExpectedBefore)
    AND (FChar = FCharBefore)
    AND (FExpectedChar = FExpectedCharBefore)
    AND (FWideChar = FWideCharBefore)
    AND (FExpectedWideChar = FExpectedWideCharBefore);
CheckFindings();
FFindingsMatch := FFindingsMatch AND FPreviewRenderingMatch;
IF (FFirstFailedScenario = 0)
    AND NOT (FResultsMatch AND FActivityMatch AND FInputsMatch AND FFindingsMatch) THEN
    FFirstFailedScenario := FScenario;
    FFailedDuringEvaluation := FEvaluateSubjects;
END_IF;
FObservationReady := TRUE;
END_METHOD

{region 'Documentation'}
(*!
<summary>Queues reset; the next bound FB call consumes it without evaluating.</summary>
*)
{endregion}
METHOD PRIVATE ResetSubjects
FText.Reset();
FWideText.Reset();
FCharacter.Reset();
FWideCharacter.Reset();
END_METHOD

